(* IEC 61131-3 sources: PLC-IsaVODE/PLC-IsaVODE/samples/plc-programs (part 3) *)

(* ---- 394-TOD_TO_STRING.ST ---- *)
FUNCTION HOUR:INT
	VAR_INPUT
		ITOD :	UDINT;
	END_VAR
	hour := UDINT_TO_INT(itod / UDINT#3600000);
END_FUNCTION

FUNCTION MINUTE:INT

	VAR_INPUT
		ITOD :	UDINT;
	END_VAR

	minute := UDINT_TO_INT((itod / UDINT#60000) - ((itod / UDINT#3600000) * UDINT#60));

END_FUNCTION

FUNCTION_BLOCK TOD_TO_STRING_Block
	VAR_INPUT
		ITOD :	UDINT;
	END_VAR

	VAR_OUTPUT
		TOD_STRING :	STRING;
	END_VAR

	VAR
		st_tmp1 :	STRING;
		st_tmp2 :	STRING;
		cur_hours :	INT;
	END_VAR

	cur_hours := hour(ITOD);
	IF cur_hours = 0 THEN
	st_tmp2 := '%01dh';
	ELSE
	st_tmp2 := '%dh';
	END_IF;

	st_tmp1 := CONCAT(INT_TO_STRING(cur_hours),INT_TO_STRING(minute(ITOD)));
	TOD_STRING := CONCAT(st_tmp1,UDINT_TO_STRING(ITOD MOD UDINT#60000 / UDINT#1000));
END_FUNCTION_BLOCK

PROGRAM program0
  VAR
    LocalVar0 : UDINT;
	LocalOUT  : STRING;
	func_block : TOD_TO_STRING_Block;
  END_VAR
	func_block.ITOD  := LocalVar0;
	func_block();
	LocalOUT := func_block.TOD_STRING;
END_PROGRAM

CONFIGURATION Config0
  RESOURCE Res0 ON PLC
    TASK task0(INTERVAL := T#20ms,PRIORITY := 0);
    PROGRAM instance0 WITH task0 : program0;
  END_RESOURCE
END_CONFIGURATION

(* ---- 396-CLICK_MODE.ST ---- *)
FUNCTION_BLOCK CLICK_MODE_Block

	VAR_INPUT
		IN :	BOOL;
		T_LONG :	TIME := T#500ms;
	END_VAR

	VAR_OUTPUT
		LONG    :   BOOL;
		SINGLE_  :	BOOL;
		DOUBLE  :	BOOL;
		TP_LONG :	BOOL;
	END_VAR

	VAR
		Timer :	TP;
		cnt :	INT;
		last :	BOOL;
	END_VAR

	timer(in := IN, PT := T_LONG);
	single := FALSE;
	double := FALSE;

	IF timer.Q THEN
		IF NOT in AND last THEN	cnt := cnt + 1; END_IF;
	ELSE
		CASE cnt OF
			1 : single := TRUE;
			2 : double := TRUE;
		END_CASE;
		cnt := 0;
	END_IF;
	last := in;
	TP_LONG := NOT timer.Q AND (NOT LONG) AND IN;
	LONG := NOT timer.Q AND in;

END_FUNCTION_BLOCK

PROGRAM program0
	VAR
		IN :	BOOL;
		T_LONG :	TIME := T#500ms;
		SINGLE_ :	BOOL;
		DOUBLE :	BOOL;
		LONG :	BOOL;
		TP_LONG :	BOOL;

		func_block : CLICK_MODE_Block;
	END_VAR
	func_block.IN := IN;
	func_block.T_LONG := T_LONG;

	func_block();
	SINGLE_  := func_block.SINGLE_;
	DOUBLE  := func_block.DOUBLE;
	LONG  := func_block.LONG;
	TP_LONG  := func_block.TP_LONG;
END_PROGRAM

CONFIGURATION Config0
	RESOURCE Res0 ON PLC
		TASK task0(INTERVAL := T#20ms,PRIORITY := 0);
		PROGRAM instance0 WITH task0 : program0;
	END_RESOURCE
END_CONFIGURATION

(* ---- 397-IP4_TO_STRING.ST ---- *)
TYPE
  oscat_STRING10             : STRING;
END_TYPE

FUNCTION _BYTE_TO_INT:INT
	VAR_INPUT
		IN :	BYTE;
	END_VAR

	_BYTE_TO_INT := USINT_TO_INT(BYTE_TO_USINT(IN));
END_FUNCTION

FUNCTION BYTE_OF_DWORD:BYTE
	VAR_INPUT
		IN :	DWORD;
		N :	BYTE;
	END_VAR
	BYTE_OF_DWORD := DWORD_TO_BYTE(SHR(in,_BYTE_TO_INT(SHL(n,3))));
END_FUNCTION

FUNCTION_BLOCK IP4_TO_STRING_Block

	VAR_INPUT
		IP4 :	DWORD;
	END_VAR

	VAR_OUTPUT
		IP4_TO_STRING :	STRING;
	END_VAR

	VAR
		s1 :	oscat_string10;
		s2 :	oscat_string10;
	END_VAR

	s1 := CONCAT(BYTE_TO_STRING(BYTE_OF_DWORD(IP4,BYTE#1)),BYTE_TO_STRING(BYTE_OF_DWORD(IP4,BYTE#0)));
	s2 := CONCAT(BYTE_TO_STRING(BYTE_OF_DWORD(IP4,BYTE#3)),BYTE_TO_STRING(BYTE_OF_DWORD(IP4,BYTE#2)));
	IP4_TO_STRING := CONCAT(s2,s1);

END_FUNCTION_BLOCK

PROGRAM program0
	VAR
		IP4 :	DWORD;
		IP4_TO_STRING :	STRING;

		func_block : IP4_TO_STRING_Block;
	END_VAR
	func_block.IP4 := IP4;

	func_block();
	IP4_TO_STRING  := func_block.IP4_TO_STRING;
END_PROGRAM

CONFIGURATION Config0

  	RESOURCE Res0 ON PLC
    	TASK task0(INTERVAL := T#20ms,PRIORITY := 0);
    	PROGRAM instance0 WITH task0 : program0;
  	END_RESOURCE

END_CONFIGURATION

(* ---- 398-SHR_4UDE.ST ---- *)
FUNCTION_BLOCK SHR_4UDE_Block

	VAR_INPUT
		SET :	BOOL;
		D0 :	BOOL;
		D3 :	BOOL;
		CLK :	BOOL;
		DN :	BOOL;
		RST :	BOOL;
	END_VAR

	VAR_OUTPUT
		Q0 :	BOOL;
		Q1 :	BOOL;
		Q2 :	BOOL;
		Q3 :	BOOL;
	END_VAR

	VAR
		trig :	R_TRIG;
	END_VAR

	trig(clk := clk);

	IF set OR rst THEN
		Q0 := NOT RST;
		Q1 := Q0;
		Q2 := Q0;
		Q3 := Q0;
	ELSIF trig.Q THEN
		IF dn THEN
			Q0 := Q1;
			Q1 := Q2;
			Q2 := Q3;
			Q3 := D3;
		ELSE
			Q3 := Q2;
			Q2 := Q1;
			Q1 := Q0;
			Q0 := D0;
		END_IF;
	END_IF;

END_FUNCTION_BLOCK

PROGRAM program0

	VAR
		SET :	BOOL;
		D0 :	BOOL;
		D3 :	BOOL;
		CLK :	BOOL;
		DN :	BOOL;
		RST :	BOOL;
		Q0 :	BOOL;
		Q1 :	BOOL;
		Q2 :	BOOL;
		Q3 :	BOOL;
		func_block : SHR_4UDE_Block;
	END_VAR
	func_block.SET  :=SET;
	func_block.D0  :=D0;
	func_block.D3  :=D3;
	func_block.CLK  :=CLK;
	func_block.DN  :=DN;
	func_block.RST  :=RST;
	func_block();
	Q0 := func_block.Q0;
	Q1 := func_block.Q1;
	Q2 := func_block.Q2;
	Q3 := func_block.Q3;

END_PROGRAM

CONFIGURATION Config0
	RESOURCE Res0 ON PLC
		TASK task0(INTERVAL := T#20ms,PRIORITY := 0);
		PROGRAM instance0 WITH task0 : program0;
	END_RESOURCE
END_CONFIGURATION

(* ---- 399-MANUAL_1.ST ---- *)
FUNCTION_BLOCK MANUAL_1_Block

	VAR_INPUT
		_IN :	BOOL;
		MAN :	BOOL;
		M_I :	BOOL;
		SET :	BOOL;
		RST :	BOOL;
	END_VAR

	VAR_OUTPUT
		Q :	BOOL;
		STATUS :	BYTE;
	END_VAR

	VAR
		S_edge :	BOOL;
		_r_edge :	BOOL;
		edge :	BOOL;
	END_VAR

	IF NOT man THEN
		Q := _IN;
		STATUS := BYTE#100;
		edge := FALSE;
	ELSIF NOT s_edge AND set THEN
		Q := TRUE;
		edge := TRUE;
		status := BYTE#101;
	ELSIF NOT _r_edge AND rst THEN
		Q := FALSE;
		edge := TRUE;
		status := BYTE#102;
	ELSIF NOT edge THEN
		Q := M_I;
		status := BYTE#103;
	END_IF;

	(* remember levels of manual signals *)
	s_edge := SET;
	_r_edge := RST;

END_FUNCTION_BLOCK

PROGRAM program0

	VAR
		_IN :	BOOL;
		MAN :	BOOL;
		M_I :	BOOL;
		SET :	BOOL;
		RST :	BOOL;

		Q :	BOOL;
		STATUS :	BYTE;

		func_block : MANUAL_1_Block;
	END_VAR
	func_block._IN := _IN;
	func_block.MAN := MAN;
	func_block.M_I := M_I;
	func_block.SET := SET;
	func_block.RST := RST;
	func_block();
	Q := func_block.Q;
	STATUS := func_block.STATUS;

END_PROGRAM

CONFIGURATION Config0

	RESOURCE Res0 ON PLC
		TASK task0(INTERVAL := T#20ms,PRIORITY := 0);
		PROGRAM instance0 WITH task0 : program0;
	END_RESOURCE

END_CONFIGURATION

(* ---- 4-COUNT_CHAR.ST ---- *)
FUNCTION_BLOCK COUNT_CHAR
	VAR_INPUT
		STR :	STRING;
		CHR :	BYTE;
	END_VAR

	VAR_OUTPUT
		COUNT_CHAR :	INT;
	END_VAR

	VAR
		I :	INT;
		pos :	INT;
	END_VAR

	I := LEN(str);
	COUNT_CHAR := 0;
	FOR pos := 1 TO I DO
		IF INT_TO_BYTE(GET_CHAR(str,pos)) = CHR THEN COUNT_CHAR := COUNT_CHAR + 1; END_IF;
	END_FOR;
END_FUNCTION_BLOCK

(* ---- 401-STRING_TO_BUFFER.ST ---- *)
TYPE
	oscat_STRING250             : STRING(250);
	oscat_arb_0_249 			  : ARRAY [0..249] 	OF BYTE;
END_TYPE

FUNCTION_BLOCK _STRING_TO_BUFFER_Block
	VAR_INPUT
		STR :	oscat_STRING250;
		POS :	INT;
		SIZE :	UINT;
	END_VAR

	VAR_OUTPUT
		_STRING_TO_BUFFER :	INT;
	END_VAR

	VAR_IN_OUT
		PT :	oscat_arb_0_249;
	END_VAR

	VAR
		i :	INT;
		end :	INT;
		x :	INT;
	END_VAR

	IF pos < 0 THEN RETURN; END_IF;
	end := MIN(pos + LEN(str), UINT_TO_INT(size)) - 1;
	x:= 1;
	FOR i := pos TO end DO
		pt[i] := INT_TO_BYTE(GET_CHAR(str,x));
		x := x + 1;
	END_FOR;

	_STRING_TO_BUFFER := i;
END_FUNCTION_BLOCK

PROGRAM program0
	VAR
	    LocalVar1 : oscat_STRING250;
        LocalVar2 : INT;
        LocalVar3 : UINT;
		LocalInOut : oscat_arb_0_249;
		LocalOUT  : INT;
		func_block : _STRING_TO_BUFFER_Block;
  	END_VAR
	func_block.STR := LocalVar1;
    func_block.POS := LocalVar2;
    func_block.SIZE := LocalVar3;
	func_block.PT := LocalInOut;
	func_block();
	LocalOUT := func_block._STRING_TO_BUFFER;
	LocalInOut := func_block.PT;
END_PROGRAM

CONFIGURATION Config0
  	RESOURCE Res0 ON PLC
    	TASK task0(INTERVAL := T#20ms,PRIORITY := 0);
    	PROGRAM instance0 WITH task0 : program0;
  	END_RESOURCE
END_CONFIGURATION

(* ---- 402-SEL2_OF_3.ST ---- *)
FUNCTION_BLOCK SEL2_OF_3_Block

	VAR_INPUT
		IN1 :	REAL;
		IN2 :	REAL;
		IN3 :	REAL;
		D :	REAL;
	END_VAR

	VAR_OUTPUT
		Y :	REAL;
		W :	INT;
		E :	BOOL;
	END_VAR

	VAR
		D12 :	BOOL;
		D23 :	BOOL;
		D31 :	BOOL;
	END_VAR

	D12 := ABS(IN1-IN2) <= D;
	D23 := ABS(IN2-IN3) <= D;
	D31 := ABS(IN3-IN1) <= D;

	IF (D12 AND D23) OR (D12 AND D31) OR (D23 AND D31) THEN
		Y := (IN1 + IN2 + IN3) * 0.333333333333;
		E := FALSE;
		W := 0;
	ELSIF D12 THEN
		Y := (In1 + IN2) * 0.5;
		E := FALSE;
		W := 3;
	ELSIF D23 THEN
		Y := (In2 + IN3) * 0.5;
		E := FALSE;
		W := 1;
	ELSIF D31 THEN
		Y := (In3 + IN1) * 0.5;
		E := FALSE;
		W := 2;
	ELSE
		E := TRUE;
		W := 4;
	END_IF;

END_FUNCTION_BLOCK

PROGRAM program0

	VAR
		IN1 :	REAL;
		IN2 :	REAL;
		IN3 :	REAL;
		D :	REAL;
		Y :	REAL;
		W :	INT;
		E :	BOOL;
		func_block : SEL2_OF_3_Block;
  	END_VAR
	func_block.IN1  :=IN1;
	func_block.IN2  :=IN2;
	func_block.IN3  :=IN3;
	func_block.D  :=D;
	func_block();
	Y := func_block.Y;
	W := func_block.W;
	E := func_block.E;

END_PROGRAM

CONFIGURATION Config0

	RESOURCE Res0 ON PLC
		TASK task0(INTERVAL := T#20ms,PRIORITY := 0);
		PROGRAM instance0 WITH task0 : program0;
	END_RESOURCE

END_CONFIGURATION

(* ---- 403-CLOG.ST ---- *)
TYPE oscat_complex :
  STRUCT
	re : REAL;
	im : REAL;
  END_STRUCT;
END_TYPE

FUNCTION ATAN2:REAL
	VAR_INPUT
		X :	REAL;
		Y :	REAL;
	END_VAR

	IF X > 0.0 THEN
		ATAN2 := ATAN(Y/X);
	ELSIF X < 0.0 THEN
		IF Y >= 0.0 THEN
			ATAN2 := ATAN(Y/X) + 3.14159265358979323846264338327950288;
		ELSE
			ATAN2 := ATAN(Y/X) - 3.14159265358979323846264338327950288;
		END_IF;
	ELSIF Y > 0.0 THEN
		ATAN2 := 1.5707963267948965580;
	ELSIF Y < 0.0 THEN
		ATAN2 := -1.5707963267948965580;
	ELSE
		ATAN2 := 0.0;
	END_IF;

END_FUNCTION

FUNCTION HYPOT:REAL
	VAR_INPUT
		X :	REAL;
		Y :	REAL;
	END_VAR

	HYPOT := SQRT(x*x + y*y);
END_FUNCTION

FUNCTION_BLOCK CLOG_Block

	VAR_INPUT
		X :	oscat_complex;
	END_VAR

	VAR_OUTPUT
		CLOG :	oscat_complex;
	END_VAR

	CLOG.re := LN(HYPOT(X.re, X.im));
	CLOG.im := ATAN2(X.im, X.re);

END_FUNCTION_BLOCK

PROGRAM program0
  VAR
    LocalVar0 : oscat_complex;
	LocalOUT  : oscat_complex;
	func_block : CLOG_Block;
  END_VAR
	func_block.X  := LocalVar0;
	func_block();
	LocalOUT := func_block.CLOG;
END_PROGRAM

CONFIGURATION Config0
  RESOURCE Res0 ON PLC
    TASK task0(INTERVAL := T#20ms,PRIORITY := 0);
    PROGRAM instance0 WITH task0 : program0;
  END_RESOURCE
END_CONFIGURATION

(* ---- 406-ELEMENT_GET.ST ---- *)
TYPE
	oscat_STRING250             : STRING;
END_TYPE

FUNCTION_BLOCK ELEMENT_GET_Block

	VAR_INPUT
		SEP :	BYTE;
		POS :	INT;
	END_VAR

	VAR_IN_OUT
		ELEMENT :	oscat_STRING250;
	END_VAR

	VAR_OUTPUT
		ELEMENT_GET :	oscat_STRING250;
	END_VAR

	VAR
		i :	INT;
		i2 :	INT;
		cnt :	INT;
		size :	INT;
	END_VAR

	cnt := 0;
	size := LEN(ELEMENT);

	FOR i := 1 TO size DO
		IF cnt = POS THEN EXIT; END_IF;
		IF INT_TO_BYTE(GET_CHAR(ELEMENT,i)) = SEP THEN cnt := cnt + 1; END_IF;
	END_FOR;

	FOR i2 := i TO size DO
		IF INT_TO_BYTE(GET_CHAR(ELEMENT,i2)) = SEP THEN EXIT; END_IF;
	END_FOR;

	IF i2 > i THEN
		ELEMENT_GET := MID(ELEMENT,i2-i,i);
	ELSE
		ELEMENT_GET := '';
	END_IF;

END_FUNCTION_BLOCK

PROGRAM program0
	VAR
		SEP :	BYTE;
		POS :	INT;
		ELEMENT :	oscat_STRING250;
		ELEMENT_GET :	oscat_STRING250;

		func_block : ELEMENT_GET_Block;
	END_VAR
	func_block.SEP    :=SEP    ;
	func_block.POS:=POS;
	func_block.ELEMENT     :=ELEMENT     ;
	func_block();
	ELEMENT    := func_block.ELEMENT    ;
	ELEMENT_GET:= func_block.ELEMENT_GET;

END_PROGRAM

CONFIGURATION Config0
  RESOURCE Res0 ON PLC
    TASK task0(INTERVAL := T#20ms,PRIORITY := 0);
    PROGRAM instance0 WITH task0 : program0;
  END_RESOURCE
END_CONFIGURATION

(* ---- 407-FILTER_MAV_DW.ST ---- *)
TYPE
  oscat_ardw_0_31             : ARRAY [0..31]   OF DWORD;
END_TYPE

FUNCTION INC1:INT

	VAR_INPUT
		X :	INT;
		N :	INT;
	END_VAR

	IF X >= N - 1 THEN
		INC1 := 0;
	ELSE
		INC1 := X + 1;
	END_IF;
END_FUNCTION

FUNCTION_BLOCK FILTER_MAV_DW

	VAR_INPUT
		X :	DWORD;
		N :	UINT;
		RST :	BOOL;
	END_VAR

	VAR_OUTPUT
		Y :	DWORD;
	END_VAR

	VAR
		init :	BOOL;
		buffer :	oscat_ardw_0_31;
		i :	INT;
		tmp :	INT;
	END_VAR

	N := MIN(N, UINT#32);

	(* startup initialisation *)
	IF NOT init OR rst OR N = UINT#0 THEN
		init := TRUE;
		tmp := UINT_TO_INT(N)-1;
		FOR i := 0 TO tmp DO
			buffer[i] := X;
		END_FOR;
		Y := X;
	ELSE
		tmp := UINT_TO_INT(N);
		i := INC1(i, tmp);
		Y := UDINT_TO_DWORD(DWORD_TO_UDINT(Y) + (DWORD_TO_UDINT(X) - DWORD_TO_UDINT(buffer[i])) / UINT_TO_UDINT(N));
		buffer[i] := X;
	END_IF;

END_FUNCTION_BLOCK

PROGRAM program0
  VAR
	X :	DWORD;
	N :	UINT;
	RST :	BOOL;

	Y :	DWORD;

	func_block : FILTER_MAV_DW;
  END_VAR
	func_block.X  := X;
	func_block.N  := N;
	func_block.RST  := RST;
	func_block();
	Y := func_block.Y;
END_PROGRAM

CONFIGURATION Config0

	RESOURCE Res0 ON PLC
		TASK task0(INTERVAL := T#20ms,PRIORITY := 0);
		PROGRAM instance0 WITH task0 : program0;
	END_RESOURCE
END_CONFIGURATION

(* ---- 409-STATUS_TO_ESR.ST ---- *)
TYPE
  oscat_esr_collect_data      : ARRAY [0..7]    OF BYTE;
END_TYPE

TYPE oscat_esr_data :
  STRUCT
	typ    : BYTE;
	adress : STRING;
	DS     : UDINT;
	TS     : TIME;
	data   : oscat_esr_collect_data;
  END_STRUCT;
END_TYPE

FUNCTION_BLOCK STATUS_TO_ESR_Block

	VAR_INPUT
		STATUS :	BYTE;
		ADRESS :	STRING;
		DT_IN :	UDINT;
		TS :	TIME;
	END_VAR

	VAR_OUTPUT
		STATUS_TO_ESR :	oscat_esr_data;
	END_VAR

	IF status < BYTE#100 THEN
		status_to_ESR.typ := BYTE#1;
	ELSIF status < BYTE#200 THEN
		status_to_ESR.typ := BYTE#2;
	ELSE
		status_to_ESR.typ := BYTE#3;
	END_IF;
	status_to_ESR.adress:= adress;
	status_to_ESR.DS := DT_in;
	status_to_ESR.TS := TS;
	status_to_ESR.data[0] := status;
END_FUNCTION_BLOCK

PROGRAM program0
	VAR
		STATUS :	BYTE;
		ADRESS :	STRING;
		DT_IN  :	UDINT;
		TS     :	TIME;
		STATUS_TO_ESR :	oscat_esr_data;

		func_block : STATUS_TO_ESR_Block;
	END_VAR
	func_block.STATUS := STATUS;
	func_block.ADRESS := ADRESS;
	func_block.DT_IN := DT_IN ;
	func_block.TS    := TS    ;

	func_block();
	STATUS_TO_ESR  := func_block.STATUS_TO_ESR;
END_PROGRAM

CONFIGURATION Config0
	RESOURCE Res0 ON PLC
		TASK task0(INTERVAL := T#20ms,PRIORITY := 0);
		PROGRAM instance0 WITH task0 : program0;
	END_RESOURCE
END_CONFIGURATION

(* ---- 410-V3_PAR.ST ---- *)
TYPE oscat_vector_3:
	STRUCT
		X : REAL;
		Y : REAL;
		Z : REAL;
	END_STRUCT;
END_TYPE

FUNCTION_BLOCK V3_ABS_Block

	VAR_INPUT
		A :	oscat_vector_3;
	END_VAR

	VAR_OUTPUT
		V3_ABS :	REAL;
	END_VAR

	V3_ABS := SQRT(A.X * A.X + A.Y * A.Y + A.Z * A.Z);

END_FUNCTION_BLOCK

FUNCTION_BLOCK V3_XPRO_Block
	VAR_INPUT
		A :	oscat_vector_3;
		B :	oscat_vector_3;
	END_VAR

	VAR_OUTPUT
		V3_XPRO :	oscat_vector_3;
	END_VAR

	V3_XPRO.X := A.Y * B.Z - A.Z * B.Y;
	V3_XPRO.Y := A.Z * B.X - A.X * B.Z;
	V3_XPRO.Z := A.X * B.Y - A.Y * B.X;

END_FUNCTION_BLOCK

FUNCTION_BLOCK V3_PAR_Block
	VAR_INPUT
		A :	oscat_vector_3;
		B :	oscat_vector_3;
	END_VAR

	VAR_OUTPUT
		V3_PAR :	BOOL;
	END_VAR

	VAR
		V3_XPRO :	V3_XPRO_Block;
		V3_ABS :	V3_ABS_Block;
	END_VAR

	V3_XPRO(A:=A,B:=B);
	V3_ABS(A:=V3_XPRO.V3_XPRO);

	V3_PAR := V3_ABS.V3_ABS = 0.0;

END_FUNCTION_BLOCK

PROGRAM program0
  	VAR
		A :	oscat_vector_3;
		B :	oscat_vector_3;
		V3_PAR :	BOOL;
		func_block : V3_PAR_Block;
  	END_VAR
	func_block.A := A;
	func_block.B := B;
	func_block();
	V3_PAR := func_block.V3_PAR;
END_PROGRAM

CONFIGURATION Config0
  RESOURCE Res0 ON PLC
    TASK task0(INTERVAL := T#20ms,PRIORITY := 0);
    PROGRAM instance0 WITH task0 : program0;
  END_RESOURCE
END_CONFIGURATION

(* ---- 411-FILTER_WAV.ST ---- *)
TYPE
  oscat_arr_0_15              : ARRAY [0..15]   OF REAL;
END_TYPE

FUNCTION INC1:INT

	VAR_INPUT
		X :	INT;
		N :	INT;
	END_VAR

	IF X >= N - 1 THEN
		INC1 := 0;
	ELSE
		INC1 := X + 1;
	END_IF;
END_FUNCTION

FUNCTION DEC1:INT

	VAR_INPUT
		X :	INT;
		N :	INT;
	END_VAR

	IF X = 0 THEN
		DEC1 := N - 1;
	ELSE
		DEC1 := X - 1;
	END_IF;

END_FUNCTION

FUNCTION_BLOCK FILTER_WAV
	VAR_INPUT
		X :	REAL;
		W :	oscat_arr_0_15;
		RST :	BOOL;
	END_VAR

	VAR_OUTPUT
		Y :	REAL;
	END_VAR

	VAR
		init :	BOOL;
		buffer :	oscat_arr_0_15;
		i :	INT;
		n :	INT;
	END_VAR

	IF NOT init OR rst THEN
		init := TRUE;
		FOR i := 0 TO 15 DO
			buffer[i] := X;
		END_FOR;
		i := 15;
		Y := X;
	ELSE
		i := INC1(i, 16);
		buffer[i] := X;
	END_IF;

	Y := 0.0;
	FOR n := 0 TO 15 DO
		Y := buffer[i] * W[n] + Y;
		i := DEC1(i, 16);
	END_FOR;
END_FUNCTION_BLOCK

PROGRAM program0
  VAR
	X :	REAL;
	W :	oscat_arr_0_15;
	RST :	BOOL;

	Y :	REAL;

	func_block : FILTER_WAV;
  END_VAR
	func_block.X  := X;
	func_block.W  := W;
	func_block.RST  := RST;
	func_block();
	Y := func_block.Y;
END_PROGRAM

CONFIGURATION Config0

	RESOURCE Res0 ON PLC
		TASK task0(INTERVAL := T#20ms,PRIORITY := 0);
		PROGRAM instance0 WITH task0 : program0;
	END_RESOURCE
END_CONFIGURATION

(* ---- 412-STRING_TO_TOD.ST ---- *)
FUNCTION_BLOCK STRING_TO_TOD_Block

  VAR_INPUT
    _TOD :	STRING;
  END_VAR

  VAR_OUTPUT
    out_STRING_TO_TOD :	UDINT;
  END_VAR

  VAR
    pos :	INT;
    i :	INT;
    tmp :	STRING;
    tmp2 :	STRING;
  END_VAR

  out_STRING_TO_TOD := UDINT#0;
  i := LEN(_TOD);
  pos :=FIND(_TOD,'#');

  IF pos>0 AND i>pos THEN
    tmp := RIGHT(_TOD,LEN(_TOD)-pos);
    pos := FIND(tmp,':');
    IF pos>1 THEN
      tmp2 := LEFT(tmp,pos-1);
      tmp := RIGHT(tmp,LEN(tmp)-pos);
      out_STRING_TO_TOD := STRING_TO_UDINT(tmp2) * UDINT#3600000;

      pos :=FIND(tmp,':');
      IF pos>1 THEN
        tmp2 := LEFT(tmp,pos-1);
        tmp := RIGHT(tmp,LEN(tmp)-pos);
        out_STRING_TO_TOD := out_STRING_TO_TOD + STRING_TO_UDINT(tmp2) * UDINT#60000;

        out_STRING_TO_TOD := out_STRING_TO_TOD + STRING_TO_UDINT(tmp) * UDINT#1000;
      END_IF;
    END_IF;
  END_IF;

END_FUNCTION_BLOCK

PROGRAM program0
  VAR
    _TOD :	STRING;
  	out_STRING_TO_TOD :	UDINT;
    func_block : STRING_TO_TOD_Block;
  END_VAR
	func_block._TOD  := _TOD;
	func_block();
	out_STRING_TO_TOD  := func_block.out_STRING_TO_TOD;
END_PROGRAM

CONFIGURATION Config0
	RESOURCE Res0 ON PLC
		TASK task0(INTERVAL := T#20ms,PRIORITY := 0);
		PROGRAM instance0 WITH task0 : program0;
	END_RESOURCE
END_CONFIGURATION

(* ---- 414-SETUP_WEEKDAYS2.ST ---- *)
TYPE
  oscat_ELEMENT_WEEKDAYS2	: ARRAY [1..7] OF STRING;
  oscat_WEEKDAYS2			: ARRAY [1..3]  OF oscat_ELEMENT_WEEKDAYS2 := [0, 0, 0];
END_TYPE

FUNCTION_BLOCK SETUP_WEEKDAYS2_Block

	VAR_IN_OUT
		WEEKDAYS2 :	oscat_WEEKDAYS2;
	END_VAR

	VAR
		init :	BOOL;
	END_VAR

	IF init THEN RETURN; END_IF;
	init := TRUE;

	WEEKDAYS2[1][01] := 'Mo';
	WEEKDAYS2[1][02] := 'Tu';
	WEEKDAYS2[1][03] := 'We';
	WEEKDAYS2[1][04] := 'Th';
	WEEKDAYS2[1][05] := 'Fr';
	WEEKDAYS2[1][06] := 'Sa';
	WEEKDAYS2[1][07] := 'Su';

	WEEKDAYS2[2][01] := 'Mo';
	WEEKDAYS2[2][02] := 'Di';
	WEEKDAYS2[2][03] := 'Mi';
	WEEKDAYS2[2][04] := 'Do';
	WEEKDAYS2[2][05] := 'Fr';
	WEEKDAYS2[2][06] := 'Sa';
	WEEKDAYS2[2][07] := 'So';

	WEEKDAYS2[3][01] := 'Lu';
	WEEKDAYS2[3][02] := 'Ma';
	WEEKDAYS2[3][03] := 'Me';
	WEEKDAYS2[3][04] := 'Je';
	WEEKDAYS2[3][05] := 'Ve';
	WEEKDAYS2[3][06] := 'Sa';
	WEEKDAYS2[3][07] := 'Di';
END_FUNCTION_BLOCK

PROGRAM program0

	VAR
		WEEKDAYS2 :	oscat_WEEKDAYS2;
		func_block : SETUP_WEEKDAYS2_Block;
	END_VAR
		func_block.WEEKDAYS2 :=WEEKDAYS2;
		func_block();
		WEEKDAYS2 := func_block.WEEKDAYS2;

END_PROGRAM

CONFIGURATION Config0

	RESOURCE Res0 ON PLC
		TASK task0(INTERVAL := T#20ms,PRIORITY := 0);
		PROGRAM instance0 WITH task0 : program0;
	END_RESOURCE

END_CONFIGURATION

(* ---- 415-STACK_16.ST ---- *)
TYPE
  oscat_ardw_0_15             : ARRAY [0..15]   OF DWORD;
END_TYPE

FUNCTION_BLOCK STACK_16_Block

	VAR_INPUT
		DIN :	DWORD;
		E :	BOOL := TRUE;
		RD :	BOOL;
		WD :	BOOL;
		RST :	BOOL;
	END_VAR

	VAR_OUTPUT
		DOUT :	DWORD;
		EMPTY :	BOOL := TRUE;
		FULL :	BOOL;
	END_VAR

	VAR
		pt :	INT;
		stack :	oscat_ardw_0_15;
	END_VAR

	IF RST THEN
		pt := 0;
		EMPTY := TRUE;
		FULL := FALSE;
		Dout := DWORD#0;
	ELSIF E THEN
		IF NOT EMPTY AND RD THEN
			pt := pt - 1;
			Dout := stack[pt];
			EMPTY := pt = 0;
			FULL := FALSE;
		END_IF;
		IF NOT FULL AND WD THEN
			stack[pt] := Din;
			pt := pt + 1;
			FULL := pt > 15;
			EMPTY := FALSE;
		END_IF;
	END_IF;

END_FUNCTION_BLOCK

PROGRAM program0
	VAR
		DIN :	DWORD;
		E :	BOOL := TRUE;
		RD :	BOOL;
		WD :	BOOL;
		RST :	BOOL;
		DOUT :	DWORD;
		EMPTY :	BOOL := TRUE;
		FULL :	BOOL;
		func_block : STACK_16_Block;
	END_VAR
		func_block.DIN  := DIN;
		func_block.E  := E;
		func_block.RD  := RD;
		func_block.WD  := WD;
		func_block.RST  := RST;
		func_block();
		DOUT := func_block.DOUT;
		EMPTY := func_block.EMPTY;
		FULL := func_block.FULL;

END_PROGRAM

CONFIGURATION Config0

	RESOURCE Res0 ON PLC
		TASK task0(INTERVAL := T#20ms,PRIORITY := 0);
		PROGRAM instance0 WITH task0 : program0;
	END_RESOURCE

END_CONFIGURATION

(* ---- 416-FILTER_MAV_W.ST ---- *)
TYPE
  oscat_FILTER_MAV_W          : ARRAY [0..31]   OF WORD;
END_TYPE

FUNCTION INC1:INT

	VAR_INPUT
		X :	INT;
		N :	INT;
	END_VAR

	IF X >= N - 1 THEN
		INC1 := 0;
	ELSE
		INC1 := X + 1;
	END_IF;
END_FUNCTION

FUNCTION_BLOCK FILTER_MAV_W
	VAR_INPUT
		X :	WORD;
		N :	UINT;
		RST :	BOOL;
	END_VAR

	VAR_OUTPUT
		Y :	WORD;
	END_VAR

	VAR
		init :	BOOL;
		buffer :	oscat_FILTER_MAV_W;
		i :	INT;
		sum :	UDINT;
		tmp :	INT;
	END_VAR

	N := MIN(N, UINT#32);

	(* startup initialisation *)
	IF NOT init OR rst OR N = UINT#0 THEN
		init := TRUE;
		tmp := UINT_TO_INT(N) - 1;
		FOR i := 1 TO tmp DO
			buffer[i] := X;
		END_FOR;
		sum := UINT_TO_UDINT(WORD_TO_UINT(Y) * N);
		Y := X;
	ELSE
		tmp := UINT_TO_INT(N);
		i := INC1(i, tmp);
		sum := sum + WORD_TO_UDINT(X) - WORD_TO_UDINT(buffer[i]);
		Y := UDINT_TO_WORD(sum / UINT_TO_UDINT(N));
		buffer[i] := X;
	END_IF;

END_FUNCTION_BLOCK

PROGRAM program0
  VAR
	X :	WORD;
	N :	UINT;
	RST :	BOOL;

	Y :	WORD;

	func_block : FILTER_MAV_W;
  END_VAR
	func_block.X  := X;
	func_block.N  := N;
	func_block.RST  := RST;
	func_block();
	Y := func_block.Y;
END_PROGRAM

CONFIGURATION Config0

	RESOURCE Res0 ON PLC
		TASK task0(INTERVAL := T#20ms,PRIORITY := 0);
		PROGRAM instance0 WITH task0 : program0;
	END_RESOURCE
END_CONFIGURATION

(* ---- 418-V3_NORM.ST ---- *)
TYPE oscat_vector_3:
	STRUCT
		X : REAL;
		Y : REAL;
		Z : REAL;
	END_STRUCT;
END_TYPE

FUNCTION_BLOCK V3_ABS_Block

	VAR_INPUT
		A :	oscat_vector_3;
	END_VAR

	VAR_OUTPUT
		V3_ABS :	REAL;
	END_VAR

	V3_ABS := SQRT(A.X * A.X + A.Y * A.Y + A.Z * A.Z);

END_FUNCTION_BLOCK

FUNCTION_BLOCK V3_SMUL_Block
	VAR_INPUT
		A :	oscat_vector_3;
		M :	REAL;
	END_VAR

	VAR_OUTPUT
		V3_SMUL :	oscat_vector_3;
	END_VAR

	V3_SMUL.X := A.X * M;
	V3_SMUL.Y := A.Y * M;
	V3_SMUL.Z := A.Z * M;
END_FUNCTION_BLOCK

FUNCTION_BLOCK V3_NORM_Block

	VAR_INPUT
		A :	oscat_vector_3;
	END_VAR

	VAR_OUTPUT
		V3_NORM :	oscat_vector_3;
	END_VAR

	VAR
		la :	REAL;
		V3_SMUL :	V3_SMUL_Block;
		V3_ABS :	V3_ABS_Block;
	END_VAR

	V3_ABS(A:=A);
	la:=V3_ABS.V3_ABS;

	IF la > 0.0 THEN
		V3_SMUL(A:=A,M:=1.0/la);
		V3_NORM:=V3_SMUL.V3_SMUL;
	ELSE
		V3_NORM.X := 0.0;
		V3_NORM.Y := 0.0;
		V3_NORM.Z := 0.0;
	END_IF;

END_FUNCTION_BLOCK

PROGRAM program0
  	VAR
		A :	oscat_vector_3;
		V3_NORM :	oscat_vector_3;
		func_block : V3_NORM_Block;
  	END_VAR
	func_block.A := A;
	func_block();
	V3_NORM := func_block.V3_NORM;
END_PROGRAM

CONFIGURATION Config0
  RESOURCE Res0 ON PLC
    TASK task0(INTERVAL := T#20ms,PRIORITY := 0);
    PROGRAM instance0 WITH task0 : program0;
  END_RESOURCE
END_CONFIGURATION

(* ---- 420-PRESSURE.ST ---- *)
FUNCTION_BLOCK PRESSURE_Block

	VAR_INPUT
		MWS :	REAL;
		TORR :	REAL;
		ATT :	REAL;
		ATM :	REAL;
		PA :	REAL;
		BAR :	REAL;
	END_VAR

	VAR_OUTPUT
		YMWS :	REAL;
		YTORR :	REAL;
		YATT :	REAL;
		YATM :	REAL;
		YPA :	REAL;
		YBAR :	REAL;
	END_VAR

	Ybar := bar +
			pa * 1.0E-5 +
			0.980665 * att +
			1.01325 * atm +
			0.001333224 * torr +
			0.0980665 * mws;
	Ymws := ybar * 10.1971621297793;
	Ytorr := ybar * 750.0615050434140;
	Yatt := ybar * 1.0197162129779;
	yatm := ybar * 0.9869232667160;
	Ypa := ybar * 100000.0;

END_FUNCTION_BLOCK

PROGRAM program0

	VAR
		MWS :	REAL;
		TORR :	REAL;
		ATT :	REAL;
		ATM :	REAL;
		PA :	REAL;
		BAR :	REAL;

		YMWS :	REAL;
		YTORR :	REAL;
		YATT :	REAL;
		YATM :	REAL;
		YPA :	REAL;
		YBAR :	REAL;
		func_block : PRESSURE_Block;
  	END_VAR
	func_block.MWS := MWS;
	func_block.TORR := TORR;
	func_block.ATT := ATT;
	func_block.ATM := ATM;
	func_block.PA := PA;
	func_block.BAR := BAR;
	func_block();
	YMWS := func_block.YMWS;
	YTORR := func_block.YTORR;
	YATT := func_block.YATT;
	YATM := func_block.YATM;
	YPA := func_block.YPA;
	YBAR := func_block.YBAR;

END_PROGRAM

CONFIGURATION Config0

  	RESOURCE Res0 ON PLC
    	TASK task0(INTERVAL := T#20ms,PRIORITY := 0);
    	PROGRAM instance0 WITH task0 : program0;
  	END_RESOURCE

END_CONFIGURATION

(* ---- 422-POLYNOM_INT.ST ---- *)
TYPE
	oscat_Polynom_ARRAY_X       : ARRAY [0..1]    OF REAL;
END_TYPE

TYPE
	oscat_Polynom_XY            : ARRAY [1..5]  OF oscat_Polynom_ARRAY_X := [0, 0, 0, 0, 0];
END_TYPE

FUNCTION_BLOCK POLYNOM_INT_Block

	VAR_INPUT
		X :	REAL;
		XY :	oscat_Polynom_XY;
	END_VAR

	VAR_INPUT
		PTS :	INT;
	END_VAR

	VAR_OUTPUT
		POLYNOM_INT :	REAL;
	END_VAR

	VAR
		XY2 :	oscat_Polynom_XY;
	END_VAR

	VAR
		I :	INT;
		J :	INT;
		J_1 :	INT;
		J_I :	INT;
		INIT :	BOOL;
	END_VAR

	pts := MIN_INT(pts, 5);

	IF (init = FALSE) THEN
		init := TRUE;

		FOR i := 1 TO pts DO
			FOR j := 0 TO 1 DO
					XY2[i][j] := XY[i][j];
			END_FOR;
		END_FOR;

		FOR i := 1 TO pts DO
			J := pts;
			WHILE (J >= i+1) DO
			j_i := j-i;
			j_1 := J-1;
			XY2[j][1] := (XY2[j][1] - XY2[j_1][1]) / (XY2[j][0] - XY2[j_i][0]);
			j := j - 1;
			END_WHILE;
		END_FOR;
	END_IF;

END_FUNCTION_BLOCK

PROGRAM program0

	VAR
		X :	REAL;
		XY :	oscat_Polynom_XY;
		PTS :	INT;

		OUT :	REAL;
		func_block : POLYNOM_INT_Block;
  	END_VAR

	func_block.X := X;
	func_block.XY := XY;
	func_block.PTS := PTS;
	func_block();
	OUT := func_block.POLYNOM_INT;

END_PROGRAM

CONFIGURATION Config0

  	RESOURCE Res0 ON PLC
    	TASK task0(INTERVAL := T#20ms,PRIORITY := 0);
    	PROGRAM instance0 WITH task0 : program0;
  	END_RESOURCE

END_CONFIGURATION

(* ---- 424-ARRAY_TREND.ST ---- *)
TYPE
	oscat_pt_ARRAY: ARRAY [1..100] OF REAL;
END_TYPE

FUNCTION BIT_OF_DWORD:BOOL
	VAR_INPUT
		IN :	DWORD;
		N :	INT;
	END_VAR
	BIT_OF_DWORD := (SHR(in,n) AND DWORD#1) > DWORD#0;
END_FUNCTION

FUNCTION EVEN:BOOL
	VAR_INPUT
		IN :	DINT;
	END_VAR
	even := NOT BIT_OF_DWORD(DINT_TO_DWORD(in),0);
END_FUNCTION

FUNCTION_BLOCK ARRAY_TREND_Block
	VAR_IN_OUT
		PT :	oscat_pt_ARRAY;
	END_VAR

	VAR_INPUT
		SIZE :	UINT;
	END_VAR

	VAR_OUTPUT
		ARRAY_TREND :	REAL;
	END_VAR

	VAR
		d :	INT;
		i :	INT;
		stop :	INT;
		stop2 :	INT;
		x :	REAL;
	END_VAR

	x := 0.0;
	stop :=LIMIT_INT(1,UINT_TO_INT(size),1000);
	stop2 := WORD_TO_INT(SHR(INT_TO_WORD(stop),1));
	IF even(INT_TO_DINT(stop)) THEN d:=0; ELSE d:=1;END_IF;

	FOR i := 1 TO stop2+d DO
		x := x - pt[i];
	END_FOR;
	FOR i := stop2+1 TO stop DO
		x := x + pt[i];
	END_FOR;
	array_trend := x / INT_TO_REAL(stop2+d);

END_FUNCTION_BLOCK

PROGRAM program0
  VAR
    LocalVar0 : oscat_pt_ARRAY;
    LocalVar1 : UINT;
	LocalOUT  : REAL;
	func_block : ARRAY_TREND_Block;
  END_VAR
	func_block.pt := LocalVar0;
	func_block.size := LocalVar1;
	func_block();
	LocalOUT := func_block.ARRAY_TREND;

END_PROGRAM

CONFIGURATION Config0
  RESOURCE Res0 ON PLC
    TASK task0(INTERVAL := T#20ms,PRIORITY := 0);
    PROGRAM instance0 WITH task0 : program0;
  END_RESOURCE
END_CONFIGURATION

(* ---- 425-SETUP_WEEKDAYS.ST ---- *)
TYPE
  oscat_ELEMENT_WEEKDAYS	: ARRAY [1..7] OF STRING;
  oscat_WEEKDAYS			: ARRAY [1..3]  OF oscat_ELEMENT_WEEKDAYS := [0, 0, 0];
END_TYPE

FUNCTION_BLOCK SETUP_WEEKDAYS

	VAR_IN_OUT
		WEEKDAYS :	oscat_WEEKDAYS;
	END_VAR

	VAR
		init :	BOOL;
	END_VAR

	IF init THEN RETURN; END_IF;
	init := TRUE;

	WEEKDAYS[1][01] := 'Monday';
	WEEKDAYS[1][02] := 'Tuesday';
	WEEKDAYS[1][03] := 'Wednesday';
	WEEKDAYS[1][04] := 'Thursday';
	WEEKDAYS[1][05] := 'Friday';
	WEEKDAYS[1][06] := 'Saturday';
	WEEKDAYS[1][07] := 'Sunday';

	WEEKDAYS[2][01] := 'Montag';
	WEEKDAYS[2][02] := 'Dienstag';
	WEEKDAYS[2][03] := 'Mittwoch';
	WEEKDAYS[2][04] := 'Donnerstag';
	WEEKDAYS[2][05] := 'Freitag';
	WEEKDAYS[2][06] := 'Samstag';
	WEEKDAYS[2][07] := 'Sonntag';

	WEEKDAYS[3][01] := 'Lundi';
	WEEKDAYS[3][02] := 'Mardi';
	WEEKDAYS[3][03] := 'Mercredi';
	WEEKDAYS[3][04] := 'Jeudi';
	WEEKDAYS[3][05] := 'Vendredi';
	WEEKDAYS[3][06] := 'Samedi';
	WEEKDAYS[3][07] := 'Dimanche';
END_FUNCTION_BLOCK

PROGRAM program0
  VAR
    WEEKDAYS :	oscat_WEEKDAYS;
	func_block : SETUP_WEEKDAYS;
  END_VAR
	func_block.WEEKDAYS  := WEEKDAYS;
	func_block();
	WEEKDAYS := func_block.WEEKDAYS;

END_PROGRAM

CONFIGURATION Config0
  RESOURCE Res0 ON PLC
    TASK task0(INTERVAL := T#20ms,PRIORITY := 0);
    PROGRAM instance0 WITH task0 : program0;
  END_RESOURCE
END_CONFIGURATION

(* ---- 426-V3_ANG.ST ---- *)
TYPE oscat_vector_3:
	STRUCT
		X : REAL;
		Y : REAL;
		Z : REAL;
	END_STRUCT;
END_TYPE

FUNCTION_BLOCK V3_ABS_Block
	VAR_INPUT
		A :	oscat_vector_3;
	END_VAR

	VAR_OUTPUT
		V3_ABS : REAL;
	END_VAR

	V3_ABS := SQRT(A.X * A.X + A.Y * A.Y + A.Z * A.Z);

END_FUNCTION_BLOCK

FUNCTION_BLOCK V3_DPRO_Block

	VAR_INPUT
		A :	oscat_vector_3;
		B :	oscat_vector_3;
	END_VAR

	VAR_OUTPUT
		V3_DPRO :	REAL;
	END_VAR

	V3_DPRO := A.X * B.X + A.Y * B.Y + A.Z * B.Z;

END_FUNCTION_BLOCK

FUNCTION_BLOCK V3_ANG_Block

	VAR_INPUT
		A :	oscat_vector_3;
		B :	oscat_vector_3;
	END_VAR

	VAR_OUTPUT
		V3_ANG :	REAL;
	END_VAR

	VAR
		d :	REAL;
		V3_ABS :	V3_ABS_Block;
		V3_DPRO :	V3_DPRO_Block;
	END_VAR

	V3_ABS(A:=A);
	d :=V3_ABS.V3_ABS;

	V3_ABS(A:=B);
	d := d * V3_ABS.V3_ABS;

	IF d > 0.0 THEN
		V3_DPRO(A:=A,B:=B);
		V3_ANG := ACOS(LIMIT(-1.0, V3_DPRO.V3_DPRO / d,1.0));
	ELSE
		V3_ANG := 0.0;

	END_IF;

END_FUNCTION_BLOCK

PROGRAM program0
  	VAR
		A :	oscat_vector_3;
		B :	oscat_vector_3;
		V3_ANG :	REAL;
		func_block : V3_ANG_Block;
  	END_VAR
	func_block.A := A;
	func_block.B := B;
	func_block();
	V3_ANG := func_block.V3_ANG;
END_PROGRAM

CONFIGURATION Config0
  RESOURCE Res0 ON PLC
    TASK task0(INTERVAL := T#20ms,PRIORITY := 0);
    PROGRAM instance0 WITH task0 : program0;
  END_RESOURCE
END_CONFIGURATION

(* ---- 427-FILL.ST ---- *)
FUNCTION_BLOCK CHR_TO_STRING_Block
	VAR_INPUT
		C :	BYTE;
	END_VAR

	VAR_OUTPUT
		CHR_TO_STRING :	STRING;
	END_VAR

	CHR_TO_STRING := BYTE_TO_STRING(C);

END_FUNCTION_BLOCK

FUNCTION BIT_OF_DWORD : BOOL
  VAR_INPUT
    IN : DWORD;
    N : INT;
  END_VAR

  BIT_OF_DWORD := (SHR(in,N) AND 16#00000001) > 0;
  (* from OSCAT library; www.oscat.de  *)
END_FUNCTION

FUNCTION_BLOCK FILL_Block
	VAR_INPUT
		C :	BYTE;
		L :	INT;
	END_VAR

	VAR_OUTPUT
		FILL :	STRING;
	END_VAR

	VAR
		N :	BYTE;
		I :	INT;
		sx :	STRING;
		CHR_TO_STRING :	CHR_TO_STRING_Block;
		FILL_tmp :	STRING;
	END_VAR

	CHR_TO_STRING(C:=c);
	Sx:=CHR_TO_STRING.CHR_TO_STRING;
	(* create string *)
	N := INT_TO_BYTE(LIMIT(0,L,80));
	(* create a string of characters to be connected to str *)
	FILL := '';
	FOR i := 1 TO 8 DO
		FILL_tmp := FILL;
		FILL := CONCAT(FILL_tmp,FILL);
		IF BIT_OF_DWORD(BYTE_TO_DWORD(N),7) THEN FILL := CONCAT(FILL,Sx); END_IF;
		N := SHL(N,1);
	END_FOR;
END_FUNCTION_BLOCK

PROGRAM program0
  VAR
	C :	BYTE;
	L :	INT;

	FILL :	STRING;

	func_block : FILL_Block;
  END_VAR
	func_block.C  :=C ;
	func_block.L  :=L ;
	func_block();
	FILL := func_block.FILL;
END_PROGRAM

CONFIGURATION Config0
  RESOURCE Res0 ON PLC
    TASK task0(INTERVAL := T#20ms,PRIORITY := 0);
    PROGRAM instance0 WITH task0 : program0;
  END_RESOURCE
END_CONFIGURATION

(* ---- 428-STACK_32.ST ---- *)
TYPE
  	oscat_ardw_0_31             : ARRAY [0..31]   OF DWORD;
END_TYPE

FUNCTION_BLOCK STACK_32_Block

	VAR_INPUT
		DIN :	DWORD;
		E :	BOOL := TRUE;
		RD :	BOOL;
		WD :	BOOL;
		RST :	BOOL;
	END_VAR

	VAR_OUTPUT
		DOUT :	DWORD;
		EMPTY :	BOOL := TRUE;
		FULL :	BOOL;
	END_VAR

	VAR
		pt :	INT;
		stack :	oscat_ardw_0_31;
	END_VAR

	IF RST THEN
		pt := 0;
		EMPTY := TRUE;
		FULL := FALSE;
		Dout := DWORD#0;
	ELSIF E THEN
		IF NOT EMPTY AND RD THEN
			(* read one element *)
			pt := pt - 1;
			Dout := stack[pt];
			EMPTY := pt = 0;
			FULL := FALSE;
		END_IF;
		IF NOT FULL AND WD THEN
			(* write one element *)
			stack[pt] := Din;
			pt := pt + 1;
			FULL := pt > 31;
			EMPTY := FALSE;
		END_IF;
	END_IF;

END_FUNCTION_BLOCK

PROGRAM program0
	VAR
		DIN :	DWORD;
		E :	BOOL := TRUE;
		RD :	BOOL;
		WD :	BOOL;
		RST :	BOOL;
		DOUT :	DWORD;
		EMPTY :	BOOL := TRUE;
		FULL :	BOOL;
		func_block : STACK_32_Block;
	END_VAR
		func_block.DIN  := DIN;
		func_block.E  := E;
		func_block.RD  := RD;
		func_block.WD  := WD;
		func_block.RST  := RST;
		func_block();
		DOUT := func_block.DOUT;
		EMPTY := func_block.EMPTY;
		FULL := func_block.FULL;

END_PROGRAM

CONFIGURATION Config0

	RESOURCE Res0 ON PLC
		TASK task0(INTERVAL := T#20ms,PRIORITY := 0);
		PROGRAM instance0 WITH task0 : program0;
	END_RESOURCE

END_CONFIGURATION

(* ---- 429-BUFFER_INSERT_NW.ST ---- *)
TYPE
  oscat_NW_BUF_LONG  : ARRAY [0..4095] OF BYTE;
END_TYPE

FUNCTION_BLOCK _BUFFER_INSERT_NW
	VAR_INPUT
		STR :	STRING;
		POS :	INT;
	END_VAR

	VAR_IN_OUT
		PT :	oscat_NW_BUF_LONG;
	END_VAR

	VAR_INPUT
		SIZE :	UINT;
	END_VAR

	VAR_OUTPUT
		_BUFFER_INSERT :	INT;
	END_VAR

	VAR
		end :	INT;
		lx :	INT;
		i :	INT;
		i2 :	INT;
		_STRING_TO_BUFFER :	_STRING_TO_BUFFER;
	END_VAR

	i := UINT_TO_INT(size) - 1;
	pos := LIMIT_INT(0,pos,i);
	lx := LEN(str);
	end := pos + lx;
	(* first move the upper part of the buffer to make space for the string *)
	i2 := i - lx;
	WHILE i >= end DO
	pt[i] := pt[i2];
	i  := i  - 1;
	i2 := i2 - 1;
	END_WHILE;

	_STRING_TO_BUFFER(str:=str, pos:=pos, size:=size, pt:=pt);
	_BUFFER_INSERT := _STRING_TO_BUFFER._STRING_TO_BUFFER;
	pt := _STRING_TO_BUFFER.pt;
END_FUNCTION_BLOCK

PROGRAM program0
  VAR
	STR :	STRING;
	POS :	INT;

	PT :	oscat_NW_BUF_LONG;

	SIZE :	UINT;

	_BUFFER_INSERT :	INT;
	func_block : _BUFFER_INSERT_NW;
  END_VAR
	func_block.STR  :=STR ;
	func_block.POS  :=POS ;
	func_block.SIZE  :=SIZE ;
	func_block.PT  :=PT ;
	func_block();
	PT := func_block.PT;
	_BUFFER_INSERT := func_block._BUFFER_INSERT;
END_PROGRAM

CONFIGURATION Config0
  RESOURCE Res0 ON PLC
    TASK task0(INTERVAL := T#20ms,PRIORITY := 0);
    PROGRAM instance0 WITH task0 : program0;
  END_RESOURCE
END_CONFIGURATION

(* ---- 430-_BUFFER_UPPERCASE_NW.ST ---- *)
TYPE
  oscat_NW_BUF_LONG  : ARRAY [0..4095] OF BYTE;
END_TYPE

FUNCTION SETUP_EXTENDED_ASCII:BOOL
	VAR_INPUT
		X :	BOOL;
	END_VAR

	SETUP_EXTENDED_ASCII := X OR TRUE;
END_FUNCTION

FUNCTION TO_UPPER:BYTE

	VAR_INPUT
		IN :	BYTE;
	END_VAR

	IF in > BYTE#96 AND in < BYTE#123 THEN
	TO_UPPER := in AND BYTE#16#DF;
	ELSIF in > BYTE#223 AND in <> BYTE#247 AND in <> BYTE#255 AND SETUP_EXTENDED_ASCII(FALSE) THEN
	TO_UPPER := in AND BYTE#16#DF;
	ELSE
	TO_UPPER := in;
	END_IF;

END_FUNCTION

FUNCTION_BLOCK _BUFFER_UPPERCASE_NW
	VAR_INPUT
		SIZE :	UINT;
	END_VAR

	VAR_OUTPUT
		_BUFFER_UPPERCASE :	BOOL;
	END_VAR

	VAR_IN_OUT
		PT :	oscat_NW_BUF_LONG;
	END_VAR

	VAR
		pos :	INT;
		size2 :	INT;
	END_VAR

	pos := 0;
	size2 := UINT_TO_INT(SIZE);

	WHILE pos < size2 DO
		PT[pos] := TO_UPPER(PT[pos]);
		pos := pos + 1;
	END_WHILE;

	_BUFFER_UPPERCASE := TRUE;

END_FUNCTION_BLOCK

PROGRAM program0
  VAR
	SIZE :	UINT;

	_BUFFER_UPPERCASE :	BOOL;

	PT :	oscat_NW_BUF_LONG;

	func_block : _BUFFER_UPPERCASE_NW;
  END_VAR
	func_block.SIZE  :=SIZE ;
	func_block.PT  :=PT ;
	func_block();
	PT := func_block.PT;
	_BUFFER_UPPERCASE := func_block._BUFFER_UPPERCASE;
END_PROGRAM

CONFIGURATION Config0
  RESOURCE Res0 ON PLC
    TASK task0(INTERVAL := T#20ms,PRIORITY := 0);
    PROGRAM instance0 WITH task0 : program0;
  END_RESOURCE
END_CONFIGURATION

(* ---- 431-SCHEDULER_2.ST ---- *)
FUNCTION_BLOCK SCHEDULER_2_Block

	VAR_INPUT
		E0 :	BOOL;
		E1 :	BOOL;
		E2 :	BOOL;
		E3 :	BOOL;
		C0 :	UINT;
		C1 :	UINT;
		C2 :	UINT;
		C3 :	UINT;
		O0 :	UINT;
		O1 :	UINT;
		O2 :	UINT;
		O3 :	UINT;
	END_VAR

	VAR_OUTPUT
		Q0 :	BOOL;
		Q1 :	BOOL;
		Q2 :	BOOL;
		Q3 :	BOOL;
	END_VAR

	VAR
		sx :	UINT;
	END_VAR

	Q0 := E0 AND (sx MOD C0 - O0 = UINT#0);
	Q1 := E1 AND (sx MOD C1 - O1 = UINT#0);
	Q2 := E2 AND (sx MOD C2 - O2 = UINT#0);
	Q3 := E3 AND (sx MOD C3 - O3 = UINT#0);

	sx := sx + UINT#1;

END_FUNCTION_BLOCK

PROGRAM program0

	VAR
		E0 :	BOOL;
		E1 :	BOOL;
		E2 :	BOOL;
		E3 :	BOOL;
		C0 :	UINT;
		C1 :	UINT;
		C2 :	UINT;
		C3 :	UINT;
		O0 :	UINT;
		O1 :	UINT;
		O2 :	UINT;
		O3 :	UINT;
		Q0 :	BOOL;
		Q1 :	BOOL;
		Q2 :	BOOL;
		Q3 :	BOOL;
		func_block : SCHEDULER_2_Block;
  	END_VAR
	func_block.E0  :=	E0;
	func_block.E1  :=	E1;
	func_block.E2  :=	E2;
	func_block.E3  :=	E3;
	func_block.C0  :=	C0;
	func_block.C1  :=	C1;
	func_block.C2  :=	C2;
	func_block.C3  :=	C3;
	func_block.O0  :=	O0;
	func_block.O1  :=	O1;
	func_block.O2  :=	O2;
	func_block.O3  :=	O3;
	func_block();
	Q0 := func_block.Q0;
	Q1 := func_block.Q1;
	Q2 := func_block.Q2;
	Q3 := func_block.Q3;

END_PROGRAM

CONFIGURATION Config0

	RESOURCE Res0 ON PLC
		TASK task0(INTERVAL := T#20ms,PRIORITY := 0);
		PROGRAM instance0 WITH task0 : program0;
	END_RESOURCE

END_CONFIGURATION

(* ---- 432-BYTE_TO_BITS.ST ---- *)
FUNCTION BIT_OF_DWORD : BOOL
  VAR_INPUT
    IN : DWORD;
    N : INT;
  END_VAR

  BIT_OF_DWORD := (SHR(in,N) AND 16#00000001) > 0;
END_FUNCTION

FUNCTION_BLOCK BYTE_TO_BITS
	VAR_INPUT
		IN :	BYTE;
	END_VAR

	VAR_OUTPUT
		B0 :	BOOL;
		B1 :	BOOL;
		B2 :	BOOL;
		B3 :	BOOL;
		B4 :	BOOL;
		B5 :	BOOL;
		B6 :	BOOL;
		B7 :	BOOL;
	END_VAR

	B0 := BIT_OF_DWORD(BYTE_TO_DWORD(IN),0); (* IN.X0 *)
	B1 := BIT_OF_DWORD(BYTE_TO_DWORD(IN),1); (* IN.X1 *)
	B2 := BIT_OF_DWORD(BYTE_TO_DWORD(IN),2); (* IN.X2 *)
	B3 := BIT_OF_DWORD(BYTE_TO_DWORD(IN),3); (* IN.X3 *)
	B4 := BIT_OF_DWORD(BYTE_TO_DWORD(IN),4); (* IN.X4 *)
	B5 := BIT_OF_DWORD(BYTE_TO_DWORD(IN),5); (* IN.X5 *)
	B6 := BIT_OF_DWORD(BYTE_TO_DWORD(IN),6); (* IN.X6 *)
	B7 := BIT_OF_DWORD(BYTE_TO_DWORD(IN),7); (* IN.X7 *)
END_FUNCTION_BLOCK

PROGRAM program0
  VAR
	LocalVar0  : BYTE;
	B0 :	BOOL;
	B1 :	BOOL;
	B2 :	BOOL;
	B3 :	BOOL;
	B4 :	BOOL;
	B5 :	BOOL;
	B6 :	BOOL;
	B7 :	BOOL;
	func_block: BYTE_TO_BITS;
  END_VAR

	func_block.IN  := LocalVar0;
	func_block();
	B0 := func_block.B0;
	B1 := func_block.B1;
	B2 := func_block.B2;
	B3 := func_block.B3;
	B4 := func_block.B4;
	B5 := func_block.B5;
	B6 := func_block.B6;
	B7 := func_block.B7;

END_PROGRAM

CONFIGURATION Config0
  RESOURCE Res0 ON PLC
    TASK task0(INTERVAL := T#20ms,PRIORITY := 0);
    PROGRAM instance0 WITH task0 : program0;
  END_RESOURCE
END_CONFIGURATION

(* ---- 433-LOG_MSG.ST ---- *)
FUNCTION_BLOCK LOG_MSG

	VAR_EXTERNAL
		LOG_CL :	us_LOG_CONTROL;
	END_VAR

	VAR
		FB_PRINT_SF :	PRINT_SF;
		idx :	INT;
	END_VAR

	IF DWORD_TO_BYTE(SHL(LOG_CL.NEW_MSG_OPTION,16)) > LOG_CL.LEVEL THEN RETURN; END_IF;
	LOG_CL.SIZE := 400;

	FB_PRINT_SF.PRINTF_DATA := LOG_CL.PRINTF;
	FB_PRINT_SF.STR 		:= LOG_CL.NEW_MSG;
	FB_PRINT_SF();
	LOG_CL.NEW_MSG	:= FB_PRINT_SF.STR;
	LOG_CL.PRINTF	:= FB_PRINT_SF.PRINTF_DATA;

	IF LOG_CL.RESET THEN
		LOG_CL.RESET := FALSE;
		LOG_CL.RING_MODE := FALSE;
		LOG_CL.IDX := 0;
		LOG_CL.UPDATE_COUNT := LOG_CL.UPDATE_COUNT + UINT#1;
	END_IF;

	IF LOG_CL.SIZE > 0 THEN
		IF LEN(LOG_CL.NEW_MSG) > 0 THEN
			IF (LOG_CL.IDX >= LOG_CL.SIZE) THEN
				LOG_CL.RING_MODE := TRUE;
				LOG_CL.IDX := 0;
			END_IF;

			LOG_CL.UPDATE_COUNT := LOG_CL.UPDATE_COUNT + UINT#1;
			LOG_CL.IDX := LOG_CL.IDX + INT#1;
			idx := LOG_CL.IDX;
			LOG_CL.MSG[idx] := LOG_CL.NEW_MSG;
			LOG_CL.MSG_OPTION[idx] := LOG_CL.NEW_MSG_OPTION;
			LOG_CL.NEW_MSG := '';
		END_IF;
	END_IF;

END_FUNCTION_BLOCK

PROGRAM program0
	VAR
		STR :	oscat_STRING80;
		LOG_MSG_R :	DWORD;
		func_block : LOG_MSG;
	END_VAR

	func_block.STR := STR;
	func_block();
	LOG_MSG_R  := func_block.LOG_MSG;
END_PROGRAM

CONFIGURATION Config0
  	RESOURCE Res0 ON PLC
    	TASK task0(INTERVAL := T#20ms,PRIORITY := 0);
    	PROGRAM instance0 WITH task0 : program0;
  	END_RESOURCE
END_CONFIGURATION

(* ---- 434-ARRAY_SDV.ST ---- *)
TYPE
	oscat_pt_ARRAY: ARRAY [1..100] OF REAL;
END_TYPE

FUNCTION_BLOCK ARRAY_VAR_Block
	VAR_IN_OUT
		PT :	oscat_pt_ARRAY;
	END_VAR

	VAR_INPUT
		SIZE :	UINT;
	END_VAR

	VAR_OUTPUT
		ARRAY_VAR :	REAL;
	END_VAR

	VAR
		i :	INT;
		stop :	INT;
		avg :	REAL;
	END_VAR

	stop :=LIMIT_INT(1,UINT_TO_INT(size),1000);
	avg := pt[1];
	FOR i := 2 TO stop DO
		avg := avg + pt[i];
	END_FOR;
	avg := avg / INT_TO_REAL(stop);

	array_var := EXPT(pt[1] - avg, 2.0);
	FOR i := 2 TO stop DO
		array_var := array_var + EXPT(pt[i] - avg, 2.0);
	END_FOR;
	array_var := array_var / INT_TO_REAL(stop-1);

END_FUNCTION_BLOCK

FUNCTION_BLOCK ARRAY_SDV_Block
	VAR_IN_OUT
		PT :	oscat_pt_ARRAY;
	END_VAR

	VAR_INPUT
		SIZE :	UINT;
	END_VAR

	VAR_OUTPUT
		ARRAY_SDV :	REAL;
	END_VAR

	VAR
		FB_array_var :	array_var_block;
	END_VAR

	FB_array_var.pt   := pt;
	FB_array_var.size := size;
	FB_array_var();
	pt := FB_array_var.pt;

	array_sdv := SQRT(FB_array_var.array_var);
END_FUNCTION_BLOCK

PROGRAM program0
  VAR
    LocalVar0 : oscat_pt_ARRAY;
    LocalVar1 : UINT;
	LocalOUT  : REAL;
	func_block : ARRAY_SDV_Block;
  END_VAR
	func_block.pt := LocalVar0;
	func_block.size := LocalVar1;
	func_block();
	LocalOUT := func_block.ARRAY_SDV;

END_PROGRAM

CONFIGURATION Config0
  RESOURCE Res0 ON PLC
    TASK task0(INTERVAL := T#20ms,PRIORITY := 0);
    PROGRAM instance0 WITH task0 : program0;
  END_RESOURCE
END_CONFIGURATION

(* ---- 435-FIFO_16.ST ---- *)
TYPE
	oscat_ardw_0_15             : ARRAY [0..15]   OF DWORD;
END_TYPE

FUNCTION INC1:INT

	VAR_INPUT
		X :	INT;
		N :	INT;
	END_VAR

	IF X >= N - 1 THEN
		INC1 := 0;
	ELSE
		INC1 := X + 1;
	END_IF;
END_FUNCTION

FUNCTION_BLOCK FIFO_16
	VAR_INPUT
		DIN :	DWORD;
		E :	BOOL := TRUE;
		RD :	BOOL;
		WD :	BOOL;
		RST :	BOOL;
	END_VAR

	VAR_OUTPUT
		DOUT :	DWORD;
		EMPTY :	BOOL := TRUE;
		FULL :	BOOL;
	END_VAR

	VAR
		fifo :	oscat_ardw_0_15;
		pr :	INT;
		pw :	INT;
	END_VAR

	IF RST THEN
		pw := pr;
		FULL := FALSE;
		EMPTY := TRUE;
		Dout := DWORD#0;
	ELSIF E THEN
		IF NOT EMPTY AND RD THEN
			Dout := fifo[pr];
			pr := INC1(pr,16);
			EMPTY := pr = pw;
			FULL := FALSE;
		END_IF;
		IF NOT FULL AND WD THEN
			fifo[pw] := Din;
			pw := INC1(pw,16);
			FULL := pw = pr;
			EMPTY := FALSE;
		END_IF;
	END_IF;
END_FUNCTION_BLOCK

PROGRAM program0
  VAR
	DIN :	DWORD;
	E   :	BOOL;
	RD  :	BOOL;
	WD  :	BOOL;
	RST :	BOOL;

	DOUT  :	DWORD;
	EMPTY :	BOOL;
	FULL  :	BOOL;

	func_block : FIFO_16;
  END_VAR
	func_block.DIN :=DIN;
	func_block.E   :=E  ;
	func_block.RD  :=RD ;
	func_block.WD  :=WD ;
	func_block.RST :=RST;
	func_block();
	DOUT := func_block.DOUT ;
	EMPTY:= func_block.EMPTY;
	FULL := func_block.FULL ;
END_PROGRAM

CONFIGURATION Config0
  RESOURCE Res0 ON PLC
    TASK task0(INTERVAL := T#20ms,PRIORITY := 0);
    PROGRAM instance0 WITH task0 : program0;
  END_RESOURCE
END_CONFIGURATION

(* ---- 437-CCOS.ST ---- *)
TYPE oscat_complex :
  STRUCT
	re : REAL;
	im : REAL;
  END_STRUCT;
END_TYPE

FUNCTION COSH:REAL
	VAR_INPUT
		X :	REAL;
	END_VAR

	VAR
		t :	REAL;
	END_VAR

	T := EXP(X);
	COSH := (1.0 / T + T) * 0.5;
END_FUNCTION

FUNCTION SINH:REAL
	VAR_INPUT
		X :	REAL;
	END_VAR

	IF ABS(x) < 2.0E-3 THEN
		SINH := X;
	ELSE
		SINH := (EXP(x) - EXP(-x)) * 0.5;
	END_IF;
END_FUNCTION

FUNCTION_BLOCK CCOSH_Block
	VAR_INPUT
		X :	oscat_complex;
	END_VAR

	VAR_OUTPUT
		CCOSH :	oscat_complex;
	END_VAR

	CCOSH.re := cosH(x.re) * COS(x.im);
	CCOSH.im := sinH(x.re) * SIN(x.im);
END_FUNCTION_BLOCK

FUNCTION_BLOCK CSET_Block
	VAR_INPUT
		RE :	REAL;
		IM :	REAL;
	END_VAR

	VAR_OUTPUT
		CSET :	oscat_complex;
	END_VAR

	CSET.re := RE;
	CSET.im := IM;
END_FUNCTION_BLOCK

FUNCTION_BLOCK CCOS_Block
	VAR_INPUT
		X :	oscat_complex;
	END_VAR

	VAR_OUTPUT
		CCOS :	oscat_complex;
	END_VAR

	VAR
		CSET :	CSET_Block;
		CCOSH :	CCOSH_Block;
	END_VAR

	CSET(RE:= -X.im,IM:=X.re);
	CCOSH(X:=CSET.CSET);
	CCOS := CCOSH.CCOSH;

END_FUNCTION_BLOCK

PROGRAM program0
  VAR
    LocalVar0 : oscat_complex;
	LocalOUT  : oscat_complex;
	func_block : CCOS_Block;
  END_VAR
	func_block.X  := LocalVar0;
	func_block();
	LocalOUT := func_block.CCOS;
END_PROGRAM

CONFIGURATION Config0
  RESOURCE Res0 ON PLC
    TASK task0(INTERVAL := T#20ms,PRIORITY := 0);
    PROGRAM instance0 WITH task0 : program0;
  END_RESOURCE
END_CONFIGURATION

(* ---- 438-FIFO_32.ST ---- *)
TYPE
	oscat_ardw_0_31             : ARRAY [0..31]   OF DWORD;
END_TYPE

FUNCTION INC1:INT

	VAR_INPUT
		X :	INT;
		N :	INT;
	END_VAR

	IF X >= N - 1 THEN
		INC1 := 0;
	ELSE
		INC1 := X + 1;
	END_IF;
END_FUNCTION

FUNCTION_BLOCK FIFO_32

	VAR_INPUT
		DIN :	DWORD;
		E :	BOOL := TRUE;
		RD :	BOOL;
		WD :	BOOL;
		RST :	BOOL;
	END_VAR

	VAR_OUTPUT
		DOUT :	DWORD;
		EMPTY :	BOOL := TRUE;
		FULL :	BOOL;
	END_VAR

	VAR
		fifo :	oscat_ardw_0_31;
		pr :	INT;
		pw :	INT;
	END_VAR

	IF RST THEN
		pw := pr;
		FULL := FALSE;
		EMPTY := TRUE;
		Dout := DWORD#0;
	ELSIF E THEN
		IF NOT EMPTY AND RD THEN
			Dout := fifo[pr];
			pr := INC1(pr,32);
			EMPTY := pr = pw;
			FULL := FALSE;
		END_IF;
		IF NOT FULL AND WD THEN
			fifo[pw] := Din;
			pw := INC1(pw,32);
			FULL := pw = pr;
			EMPTY := FALSE;
		END_IF;
	END_IF;

END_FUNCTION_BLOCK

PROGRAM program0
  VAR
	DIN :	DWORD;
	E   :	BOOL;
	RD  :	BOOL;
	WD  :	BOOL;
	RST :	BOOL;

	DOUT  :	DWORD;
	EMPTY :	BOOL;
	FULL  :	BOOL;

	func_block : FIFO_32;
  END_VAR
	func_block.DIN :=DIN;
	func_block.E   :=E  ;
	func_block.RD  :=RD ;
	func_block.WD  :=WD ;
	func_block.RST :=RST;
	func_block();
	DOUT := func_block.DOUT ;
	EMPTY:= func_block.EMPTY;
	FULL := func_block.FULL ;
END_PROGRAM

CONFIGURATION Config0
  RESOURCE Res0 ON PLC
    TASK task0(INTERVAL := T#20ms,PRIORITY := 0);
    PROGRAM instance0 WITH task0 : program0;
  END_RESOURCE
END_CONFIGURATION

(* ---- 439-ALARM_2.ST ---- *)
FUNCTION_BLOCK ALARM_2
	VAR_INPUT
		X :	REAL;
		LO_1 :	REAL;
		HI_1 :	REAL;
		LO_2 :	REAL;
		HI_2 :	REAL;
		HYS :	REAL;
	END_VAR

	VAR_OUTPUT
		Q1_LO :	BOOL;
		Q1_HI :	BOOL;
		Q2_LO :	BOOL;
		Q2_HI :	BOOL;
	END_VAR

	VAR
		tmp :	REAL;
	END_VAR

	tmp := X - Hys * 0.5;
	IF tmp > LO_1 THEN Q1_LO := FALSE; END_IF;
	IF tmp > LO_2 THEN Q2_LO := FALSE; END_IF;
	IF tmp > HI_1 THEN Q1_HI := TRUE; END_IF;
	IF tmp > HI_2 THEN Q2_HI := TRUE; END_IF;
	tmp := tmp + hys;
	IF tmp < LO_1 THEN Q1_LO := TRUE; END_IF;
	IF tmp < LO_2 THEN Q2_LO := TRUE; END_IF;
	IF tmp < HI_1 THEN Q1_HI := FALSE; END_IF;
	IF tmp < HI_2 THEN Q2_HI := FALSE; END_IF;

END_FUNCTION_BLOCK

PROGRAM program0
	VAR
	    LocalVar0 : REAL;
		LocalVar1 : REAL;
		LocalVar2 : REAL;
		LocalVar3 : REAL;
		LocalVar4 : REAL;
		LocalVar5 : REAL;
		LocalOUT1  : BOOL;
		LocalOUT2  : BOOL;
		LocalOUT3  : BOOL;
		LocalOUT4  : BOOL;
		func_block : ALARM_2;
  	END_VAR
	func_block.X := LocalVar0;
	func_block.LO_1 := LocalVar1;
	func_block.HI_1 := LocalVar2;
	func_block.LO_2 := LocalVar3;
	func_block.HI_2 := LocalVar4;
	func_block.HYS := LocalVar5;
	func_block();
	LocalOUT1 := func_block.Q1_LO;
	LocalOUT2 := func_block.Q1_HI;
	LocalOUT3 := func_block.Q2_LO;
	LocalOUT4 := func_block.Q2_HI;
END_PROGRAM

CONFIGURATION Config0
  	RESOURCE Res0 ON PLC
    	TASK task0(INTERVAL := T#20ms,PRIORITY := 0);
    	PROGRAM instance0 WITH task0 : program0;
  	END_RESOURCE
END_CONFIGURATION

(* ---- 440-DRIVER_4C.ST ---- *)
TYPE
  oscat_DRIVER_4C 			  : ARRAY [1..7] 	OF BYTE;
END_TYPE
FUNCTION_BLOCK DRIVER_4C

	VAR_INPUT
		IN :	BOOL;
		RST :	BOOL;
		TIMEOUT :	TIME;
		SX :	oscat_DRIVER_4C;
	END_VAR

	VAR_OUTPUT
		SN :	INT;
		Q0 :	BOOL;
		Q1 :	BOOL;
		Q2 :	BOOL;
		Q3 :	BOOL;
	END_VAR

	VAR
		off :	TON;
		edge :	BOOL;
	END_VAR

	IF RST OR off.Q THEN
		SN := 0;
	ELSIF IN AND NOT edge THEN
		SN := SN + 1;
		IF SN > 7 OR SX[SN] = BYTE#0 THEN SN := 0; END_IF;
	END_IF;
	edge := in;
	IF SN > 0 THEN
		Q0 := (SX[SN] AND BYTE#1) > BYTE#0;
		Q1 := (SX[SN] AND BYTE#2) > BYTE#0;
		Q2 := (SX[SN] AND BYTE#4) > BYTE#0;
		Q3 := (SX[SN] AND BYTE#8) > BYTE#0;
	ELSE
		Q0 := FALSE;
		Q1 := FALSE;
		Q2 := FALSE;
		Q3 := FALSE;
	END_IF;

	IF timeout > t#0s THEN off(in := SN > 0, PT := Timeout); END_IF;

END_FUNCTION_BLOCK

PROGRAM program0
  VAR
	IN      :	BOOL;
	RST     :	BOOL;
	TIMEOUT :	TIME;
	SX      :	oscat_DRIVER_4C;

	SN :	INT;
	Q0 :	BOOL;
	Q1 :	BOOL;
	Q2 :	BOOL;
	Q3 :	BOOL;

	func_block : DRIVER_4C;
  END_VAR
	func_block.IN       :=IN      ;
	func_block.RST      :=RST     ;
	func_block.TIMEOUT  :=TIMEOUT ;
	func_block.SX       :=SX      ;
	func_block();
	SN := func_block.SN;
	Q0 := func_block.Q0;
	Q1 := func_block.Q1;
	Q2 := func_block.Q2;
	Q3 := func_block.Q3;
END_PROGRAM

CONFIGURATION Config0
  RESOURCE Res0 ON PLC
    TASK task0(INTERVAL := T#20ms,PRIORITY := 0);
    PROGRAM instance0 WITH task0 : program0;
  END_RESOURCE
END_CONFIGURATION

(* ---- 441-COUNT_DR.ST ---- *)
FUNCTION_BLOCK COUNT_DR
	VAR_INPUT
		SET :	BOOL;
		IN :	DWORD;
		UP :	BOOL;
		DN :	BOOL;
		STEPP :	DWORD := DWORD#1;
		MX :	DWORD := DWORD#16#FFFF_FFFF;
		RST :	BOOL;
	END_VAR

	VAR_OUTPUT
		CNT :	DWORD;
	END_VAR

	VAR
		CNT2 :	UDINT;
		STEPP2 :	UDINT;
		MX2 :	UDINT;
		last_up :	BOOL;
		last_dn :	BOOL;
	END_VAR

	STEPP2 := DWORD_TO_UDINT(STEPP);
	MX2   := DWORD_TO_UDINT(MX);
	CNT2  := DWORD_TO_UDINT(CNT);

	IF rst THEN
		CNT2 := UDINT#0;
	ELSIF set THEN
		CNT2 := LIMIT(UDINT#0,DWORD_TO_UDINT(in),mx2);
	ELSIF up AND NOT last_up THEN
		IF STEPP2 > MX2 - CNT2 THEN
			CNT2 := CNT2 - MX2 + STEPP2 - UDINT#1;
		ELSE
			CNT2 := CNT2 + STEPP2;
		END_IF;
	ELSIF dn AND NOT last_dn THEN
		IF STEPP2 > CNT2 THEN
			CNT2 := CNT2 - STEPP2 + MX2 + UDINT#1;
		ELSE
			CNT2 := CNT2 - STEPP2;
		END_IF;
	END_IF;
	last_up := up;
	last_dn := dn;
	CNT := UDINT_TO_DWORD(CNT2);
END_FUNCTION_BLOCK

PROGRAM program0
  VAR
	SET :	BOOL;
	IN :	DWORD;
	UP :	BOOL;
	DN :	BOOL;
	STEPP :	DWORD;
	MX :	DWORD;
	RST :	BOOL;

	CNT :	DWORD;
	func_block : COUNT_DR;
  END_VAR
	func_block.SET  :=SET  ;
	func_block.IN   :=IN   ;
	func_block.UP   :=UP   ;
	func_block.DN   :=DN   ;
	func_block.STEPP :=STEPP ;
	func_block.MX   :=MX   ;
	func_block.RST  :=RST  ;

	func_block();
	CNT := func_block.CNT;
END_PROGRAM

CONFIGURATION Config0
  RESOURCE Res0 ON PLC
    TASK task0(INTERVAL := T#20ms,PRIORITY := 0);
    PROGRAM instance0 WITH task0 : program0;
  END_RESOURCE
END_CONFIGURATION

(* ---- 442-BUFFER_SEARCH.ST ---- *)
TYPE
	oscat_arb_0_249 			  : ARRAY [0..249] 	OF BYTE;
END_TYPE

FUNCTION_BLOCK BUFFER_SEARCH_Block
	VAR_INPUT
		SIZE :	UINT;
		STR :	STRING;
		POS :	INT;
		IGN :	BOOL;
	END_VAR

	VAR_IN_OUT
		PT :	oscat_arb_0_249;
	END_VAR

	VAR_OUTPUT
		BUFFER_SEARCH :	INT;
	END_VAR

	VAR
		i :	INT;
		end :	INT;
		k :	INT;
		k2 :	INT;
		lx :	INT;
		char :	BYTE;
		chx :	BYTE;
	END_VAR

	lx := LEN(str);
	IF pos >= 0 AND lx > 0 THEN
		end := UINT_TO_INT(size) - lx;
		lx := lx - 1;
		FOR i := pos TO end DO
			FOR k := 0 TO lx DO
				char := INT_TO_BYTE(GET_CHAR(str,k + 1));
				k2 := i + k;
				IF IGN THEN
					chx := TO_UPPER(pt[k2]);
				ELSE
					chx := pt[k2];
				END_IF;
				IF char <> chx THEN EXIT; END_IF;
			END_FOR;
			IF k > lx THEN
				BUFFER_SEARCH := i;
				RETURN;
			END_IF;
		END_FOR;
	END_IF;
	BUFFER_SEARCH := -1;
END_FUNCTION_BLOCK

PROGRAM program0
  VAR
    LocalVar0 : UINT;
    LocalVar1 : STRING;
	LocalVar2 : INT;
	LocalVar3 : BOOL;
	LocalVar4 : oscat_arb_0_249;
	LocalOUT  : INT;
	func_block : BUFFER_COMP_Block;
  END_VAR
	func_block.SIZE  := LocalVar0;
	func_block.STR  := LocalVar1;
	func_block.POS   := LocalVar2;
	func_block.IGN  := LocalVar3;
	func_block.PT := LocalVar4;
	func_block();
	LocalOUT := func_block.BUFFER_COMP;
	LocalVar4 := func_block.PT;

END_PROGRAM

CONFIGURATION Config0
  RESOURCE Res0 ON PLC
    TASK task0(INTERVAL := T#20ms,PRIORITY := 0);
    PROGRAM instance0 WITH task0 : program0;
  END_RESOURCE
END_CONFIGURATION

(* ---- 445-COUNT_BR.ST ---- *)
FUNCTION _BYTE_TO_INT:INT
	VAR_INPUT
		IN :	BYTE;
	END_VAR

	_BYTE_TO_INT := USINT_TO_INT(BYTE_TO_USINT(IN));

END_FUNCTION

FUNCTION INC:INT
	VAR_INPUT
		X :	INT;
		D :	INT;
		M :	INT;
	END_VAR

	inc := (X + D + M + 1) MOD (M + 1);
END_FUNCTION

FUNCTION_BLOCK COUNT_BR
	VAR_INPUT
		SET :	BOOL;
		IN :	BYTE;
		UP :	BOOL;
		DN :	BOOL;
		STEPP :	BYTE := BYTE#1;
		MX :	BYTE := BYTE#255;
		RST :	BOOL;
	END_VAR
	VAR_OUTPUT
		CNT :	BYTE;
	END_VAR

	VAR
		last_up :	BOOL;
		last_dn :	BOOL;
	END_VAR

	IF rst THEN
		cnt := BYTE#0;
	ELSIF set THEN
		cnt := INT_TO_BYTE(LIMIT(0,_BYTE_TO_INT(in),_BYTE_TO_INT(mx)));
	ELSIF up AND NOT last_up THEN
		cnt := INT_TO_BYTE(inc(_BYTE_TO_INT(cnt),_BYTE_TO_INT(stepP),_BYTE_TO_INT(mx)));
	ELSIF dn AND NOT last_dn THEN
		cnt := INT_TO_BYTE(inc(_BYTE_TO_INT(cnt),_BYTE_TO_INT(stepP) * -1,_BYTE_TO_INT(mx)));
	END_IF;
	last_up := up;
	last_dn := dn;
END_FUNCTION_BLOCK

PROGRAM program0
  VAR
	SET :	BOOL;
	IN :	BYTE;
	UP :	BOOL;
	DN :	BOOL;
	STEPP:	BYTE;
	MX :	BYTE;
	RST :	BOOL;

	CNT :	BYTE;
	func_block : COUNT_BR;
  END_VAR
	func_block.SET  :=SET  ;
	func_block.IN   :=IN   ;
	func_block.UP   :=UP   ;
	func_block.DN   :=DN   ;
	func_block.STEPP :=STEPP ;
	func_block.MX   :=MX   ;
	func_block.RST  :=RST  ;

	func_block();
	CNT := func_block.CNT;
END_PROGRAM

CONFIGURATION Config0
  RESOURCE Res0 ON PLC
    TASK task0(INTERVAL := T#20ms,PRIORITY := 0);
    PROGRAM instance0 WITH task0 : program0;
  END_RESOURCE
END_CONFIGURATION

(* ---- 446-RC4_CRYPT_STREAM.ST ---- *)
FUNCTION_BLOCK RC4_CRYPT_STREAM

	VAR_IN_OUT
		MODE :	INT;
		KEY :	oscat_STRING40;
		BUF :	oscat_aB0_63;
		SIZE :	UDINT;
	END_VAR

	VAR_OUTPUT
		POS :	UDINT;
	END_VAR

	VAR
		sbox :	oscat_aB0_255;
		skey :	oscat_aB0_255;
		a :	INT;
		b :	INT;
		c :	INT;
		d :	USINT;
		e :	USINT;
		end :	UDINT;
		v :	BYTE;
		v_tmp :	INT;
		CODE :	CODE;
	END_VAR

	CASE MODE OF

	1:
		b := LEN(KEY) - 1;
		IF b < 0 OR SIZE < UDINT#1 THEN
			MODE := 3;
			RETURN;
		END_IF;

		FOR a := 0 TO b DO
			CODE(STR:=KEY,POS:=a + 1);
			skey[a] := CODE.CODE;
			sbox[a] := INT_TO_BYTE(a);
		END_FOR;

		c := 0;
		FOR a := b + 1 TO 255 DO
			skey[a] := skey[c];
			sbox[a] := INT_TO_BYTE(a);
			c := c + 1;
			IF c > b THEN c := 0; END_IF;
		END_FOR;

		d := USINT#0;
		FOR a := 0 TO 255 DO
			d := d + BYTE_TO_USINT(sbox[a]) + BYTE_TO_USINT(skey[a]);
			v := sbox[a];
			sbox[a] := sbox[d];
			sbox[d] := v;
		END_FOR;

		POS := UDINT#0;
		end := SIZE;
		SIZE := MIN(UDINT#64,end);
		d := USINT#0;
		e := USINT#0;
		MODE := 2;

	2:

		b := UDINT_TO_INT(SIZE) - 1;
		FOR a := 0 TO b DO
			d := d + USINT#1;
			e := e + BYTE_TO_USINT(sbox[d]);
			v := sbox[d];
			sbox[d] := sbox[e];
			sbox[e] := v;
			v := USINT_TO_BYTE(BYTE_TO_USINT(sbox[d]) + BYTE_TO_USINT(sbox[e]));
			v_tmp := _BYTE_TO_INT(v);
			BUF[a] :=BUF[a] XOR sbox[v_tmp];
		END_FOR;

		POS := POS + SIZE;
		SIZE := MIN(UDINT#64,end - POS);

		IF SIZE = UDINT#0 THEN
			MODE := 3;
		END_IF;
	END_CASE;

END_FUNCTION_BLOCK

(* ---- 448-T_PLC_US.ST ---- *)
FUNCTION_BLOCK T_PLC_US_Block

	VAR_OUTPUT
		T_PLC_US :	UDINT;
	END_VAR

	VAR_EXTERNAL
		PLC_TICKS_PER_SEC :	INT;
		PLC_SYS_TICK_CNT :	DINT;
	END_VAR

	VAR
		debug :	BOOL;
		N :	INT;
		Offset :	UDINT;
		temp :	DWORD := DWORD#1;
		mode :	BOOL;
		faktor :	UDINT;
		init :	BOOL;
		v_plc_ticks_per_sec :	UDINT;
		base :	UDINT := UDINT#1000000;
	END_VAR

	IF init = FALSE THEN
		v_plc_ticks_per_sec := INT_TO_UDINT(PLC_TICKS_PER_SEC);
		IF v_plc_ticks_per_sec = UDINT#1024 THEN
			faktor := UDINT#1000;
			mode := FALSE;
		ELSIF v_plc_ticks_per_sec > UDINT#0 THEN
			IF v_plc_ticks_per_sec <= base THEN
				faktor := base / v_plc_ticks_per_sec;
				mode := FALSE;
			ELSE
				faktor := v_plc_ticks_per_sec / base;
				mode := TRUE;
			END_IF;
		ELSE
			faktor := UDINT#1;
		END_IF;
		init := TRUE;
	END_IF;

	IF mode THEN
		T_PLC_US := DINT_TO_UDINT(PLC_SYS_TICK_CNT) / faktor;
	ELSE
		T_PLC_US := DINT_TO_UDINT(PLC_SYS_TICK_CNT) * faktor;
	END_IF;

	IF debug THEN
		T_PLC_US := (DWORD_TO_UDINT(SHL(UDINT_TO_DWORD(T_PLC_US),N) OR SHL(temp,N)) - UDINT#1) + Offset;
	END_IF;

END_FUNCTION_BLOCK

PROGRAM program0

	VAR
		T_PLC_US  : UDINT;
		func_block : T_PLC_US_Block;
	END_VAR
		func_block();
		T_PLC_US := func_block.T_PLC_US;

END_PROGRAM

CONFIGURATION Config0

	VAR_GLOBAL
		PLC_TICKS_PER_SEC :	INT;
		PLC_SYS_TICK_CNT :	DINT;
	END_VAR

	RESOURCE Res0 ON PLC
		TASK task0(INTERVAL := T#20ms,PRIORITY := 0);
		PROGRAM instance0 WITH task0 : program0;
	END_RESOURCE

END_CONFIGURATION

(* ---- 449-REAL_TO_STRF.ST ---- *)
FUNCTION EXP10 : REAL

	VAR_INPUT
		x : REAL;
	END_VAR

	exp10 := EXP(X * 2.30258509299405);

END_FUNCTION

FUNCTION _REAL_TO_DINT:DINT
	VAR_INPUT
		X :	REAL;
	END_VAR

	IF REAL_TO_DINT(0.5) = DINT#1 THEN
		_REAL_TO_DINT := REAL_TO_DINT(x);
		RETURN;
	END_IF;

	IF X > 0.0 THEN
		_REAL_TO_DINT := REAL_TO_DINT(x+0.5);
	ELSIF X < 0.0 THEN
		_REAL_TO_DINT := REAL_TO_DINT(x-0.5);
	ELSE
		_REAL_TO_DINT := DINT#0;
	END_IF;
END_FUNCTION

FUNCTION_BLOCK REAL_TO_STRF_Block

	VAR_INPUT
		IN :	REAL;
		N :	INT;
		D :	STRING;
	END_VAR

	VAR_OUTPUT
		REAL_TO_STRF :	STRING;
	END_VAR

	VAR
		st_tmp : STRING;
		i :	INT;
	END_VAR

	N := LIMIT(0,N,7);
	REAL_TO_STRF := DINT_TO_STRING(_REAL_TO_DINT(ABS(in) * EXP10(INT_TO_REAL(N))));
	FOR i := LEN(REAL_TO_STRF) TO N DO
		st_tmp := REAL_TO_STRF;
		REAL_TO_STRF := CONCAT('0', st_tmp);
	END_FOR;
	IF n > 0 THEN REAL_TO_STRF := INSERT(REAL_TO_STRF, D, LEN(REAL_TO_STRF) - N); END_IF;
	IF in < 0.0 THEN st_tmp := REAL_TO_STRF; REAL_TO_STRF := CONCAT('-', st_tmp); END_IF;

END_FUNCTION_BLOCK

PROGRAM program0

	VAR
		IN :	REAL;
		N :	INT;
		D :	STRING;

        REAL_TO_STRF :	STRING;
		func_block : REAL_TO_STRF_Block;
	END_VAR
		func_block.IN := IN;
		func_block.N := N;
		func_block.D := D;
		func_block();
		REAL_TO_STRF := func_block.REAL_TO_STRF;

END_PROGRAM

CONFIGURATION Config0

	RESOURCE Res0 ON PLC
		TASK task0(INTERVAL := T#20ms,PRIORITY := 0);
		PROGRAM instance0 WITH task0 : program0;
	END_RESOURCE

END_CONFIGURATION

(* ---- 452-MESSAGE_4R.ST ---- *)
FUNCTION INC1:INT

	VAR_INPUT
		X :	INT;
		N :	INT;
	END_VAR

	IF X >= N - 1 THEN
		INC1 := 0;
	ELSE
		INC1 := X + 1;
	END_IF;
END_FUNCTION

FUNCTION_BLOCK MESSAGE_4R_Block

	VAR_INPUT
		M0 :	STRING;
		M1 :	STRING;
		M2 :	STRING;
		M3 :	STRING;
		MM :	INT := 3;
		ENQ :	BOOL := TRUE;
		CLK :	BOOL := TRUE;
		T1 :	TIME := T#3s;
	END_VAR

	VAR_OUTPUT
		MX :	STRING;
		MN :	INT;
		TR :	BOOL;
	END_VAR

	VAR
		timer :	TON;
		edge :	BOOL;
	END_VAR

	TR := FALSE;
	IF ENQ THEN
		IF (NOT edge AND clk) OR timer.q THEN
				MN := INC1(MN, MM);
				TR := TRUE;
				timer(in := FALSE);
				CASE MN OF
					0 : MX := M0;
					1 : MX := M1;
					2 : MX := M2;
					3 : MX := M3;
				END_CASE;
		END_IF;
		edge := clk;
		timer( in := CLK, pt := T1);
	ELSE
		MX := '';
		MN := 0;
	END_IF;

END_FUNCTION_BLOCK

PROGRAM program0

	VAR
		M0 :	STRING;
		M1 :	STRING;
		M2 :	STRING;
		M3 :	STRING;
		MM :	INT;
		ENQ :	BOOL;
		CLK :	BOOL;
		T1 :	TIME;

		MX :	STRING;
		MN :	INT;
		TR :	BOOL;

		func_block : MESSAGE_4R_Block;
	END_VAR

	func_block.M0 := M0;
	func_block.M1 := M1;
	func_block.M2 := M2;
	func_block.M3 := M3;
	func_block.MM := MM;
	func_block.ENQ := ENQ;
	func_block.CLK := CLK;
	func_block.T1 := T1;

	func_block();

	MX := func_block.MX;
	MN := func_block.MN;
	TR := func_block.TR;

END_PROGRAM

CONFIGURATION Config0

	RESOURCE Res0 ON PLC
		TASK task0(INTERVAL := T#20ms,PRIORITY := 0);
		PROGRAM instance0 WITH task0 : program0;
	END_RESOURCE

END_CONFIGURATION

(* ---- 453-BASE64_DECODE_STREAM.ST ---- *)
TYPE
  oscat_aB0_47	: ARRAY [0..47]	OF BYTE;
  oscat_aB0_63	: ARRAY [0..63]	OF BYTE;
END_TYPE

FUNCTION_BLOCK BASE64_DECODE_STREAM
	VAR_IN_OUT
		BUF1 :	oscat_aB0_63;
		BUF2 :	oscat_aB0_47;
	END_VAR

	VAR_INPUT
		SIZE1 :	INT;
	END_VAR

	VAR_OUTPUT
		SIZE2 :	INT;
	END_VAR

	VAR
		a :	INT;
		b :	WORD;
		o :	INT;
		off :	INT;
		i1 :	INT;
		i2 :	INT;
		c :	INT;
	END_VAR

	IF SIZE1 <= 0 THEN SIZE2 := 0; RETURN; END_IF;
	c := SIZE1 - 1;
	i2 := 0;
	a := 0;
	b := WORD#0;
	FOR i1 := 0 TO c DO
		o := BYTE_TO_INT(BUF1[i1]);
		IF o = 61  (* = *) THEN EXIT;
		ELSIF o > 96 (* a-z *) THEN off := 71;
		ELSIF o > 64 (* A-Z *) THEN off := 65;
		ELSIF o > 47 (* 0-9 *) THEN off := -4;
		ELSIF o = 43 (* + *) THEN off := -19;
		ELSIF o = 47 (* / *) THEN off := -16;
		END_IF;
		b := SHL(b,6) OR INT_TO_WORD(o - off);
		a := a + 6;
		IF a >= 8 THEN
			a := a - 8;
			BUF2[i2] := WORD_TO_BYTE(SHR(b,a));
			i2 := i2 + 1;
			b := b AND NOT SHL(WORD#16#FFFF,a);
		END_IF;
	END_FOR;
	SIZE2 := i2;
END_FUNCTION_BLOCK

PROGRAM program0
  VAR
	BUF1  :	oscat_aB0_63;
	BUF2  :	oscat_aB0_47;

	SIZE1 :	INT;

	SIZE2 :	INT;
	func_block : BASE64_DECODE_STREAM;
  END_VAR
	func_block.BUF1 :=BUF1 ;
	func_block.BUF2 :=BUF2 ;
	func_block.SIZE1:=SIZE1;
	func_block();
	BUF1 := func_block.BUF1;
	BUF2 := func_block.BUF2;
	SIZE2 := func_block.SIZE2;
END_PROGRAM

CONFIGURATION Config0
  RESOURCE Res0 ON PLC
    TASK task0(INTERVAL := T#20ms,PRIORITY := 0);
    PROGRAM instance0 WITH task0 : program0;
  END_RESOURCE
END_CONFIGURATION

(* ---- 456-SHR_8UDE.ST ---- *)
FUNCTION_BLOCK SHR_8UDE_Block

	VAR_INPUT
		SET :	BOOL;
		D0 :	BOOL;
		D7 :	BOOL;
		CLK :	BOOL;
		DN :	BOOL;
		RST :	BOOL;
	END_VAR

	VAR_OUTPUT
		Q0 :	BOOL;
		Q1 :	BOOL;
		Q2 :	BOOL;
		Q3 :	BOOL;
		Q4 :	BOOL;
		Q5 :	BOOL;
		Q6 :	BOOL;
		Q7 :	BOOL;
	END_VAR

	VAR
		trig :	R_TRIG;
	END_VAR

	trig(clk := clk);

	IF set OR rst THEN
		Q0 := NOT RST;
		Q1 := Q0;
		Q2 := Q0;
		Q3 := Q0;
		Q4 := Q0;
		Q5 := Q0;
		Q6 := Q0;
		Q7 := Q0;
	ELSIF trig.Q THEN
		IF dn THEN
			Q0 := Q1;
			Q1 := Q2;
			Q2 := Q3;
			Q3 := Q4;
			Q4 := Q5;
			Q5 := Q6;
			Q6 := Q7;
			Q7 := D7;
		ELSE
			Q7 := Q6;
			Q6 := Q5;
			Q5 := Q4;
			Q4 := Q3;
			Q3 := Q2;
			Q2 := Q1;
			Q1 := Q0;
			Q0 := D0;
		END_IF;
	END_IF;

END_FUNCTION_BLOCK

PROGRAM program0
	VAR
		SET :	BOOL;
		D0 :	BOOL;
		D7 :	BOOL;
		CLK :	BOOL;
		DN :	BOOL;
		RST :	BOOL;
		Q0 :	BOOL;
		Q1 :	BOOL;
		Q2 :	BOOL;
		Q3 :	BOOL;
		Q4 :	BOOL;
		Q5 :	BOOL;
		Q6 :	BOOL;
		Q7 :	BOOL;
		func_block : SHR_8UDE_Block;
  	END_VAR
	func_block.SET  :=SET;
	func_block.D0  :=D0;
	func_block.D7  :=D7;
	func_block.CLK  :=CLK;
	func_block.DN  :=DN;
	func_block.RST  :=RST;
	func_block();
	Q0  := func_block.Q0;
	Q1  := func_block.Q1;
	Q2  := func_block.Q2;
	Q3  := func_block.Q3;
	Q4  := func_block.Q4;
	Q5  := func_block.Q5;
	Q6  := func_block.Q6;
	Q7  := func_block.Q7;
END_PROGRAM

CONFIGURATION Config0
	RESOURCE Res0 ON PLC
		TASK task0(INTERVAL := T#20ms,PRIORITY := 0);
		PROGRAM instance0 WITH task0 : program0;
	END_RESOURCE
END_CONFIGURATION

(* ---- 457-TELNET_LOG.ST ---- *)
FUNCTION_BLOCK TELNET_LOG

	VAR_INPUT
		ENABLE :	BOOL;
		OPTION :	BYTE := BYTE#2#1000_1100;
		PORT :	WORD := WORD#23;
	END_VAR

	VAR_OUTPUT
		READY :	BOOL;
	END_VAR

	VAR_IN_OUT
		IP_C :	oscat_IP_C;
		S_BUF :	oscat_NETWORK_BUFFER;
		LOG_CL :	us_LOG_CONTROL;
	END_VAR

	VAR
		TELNET_PRINT :	TELNET_PRINT;
		done :	BOOL;
		init :	BOOL;
		watchdog :	TON;
		ci :	INT;
		pi :	INT;
		pi_last :	INT;
		send :	BOOL;
	END_VAR

	IF NOT init THEN
		init := TRUE;
		IF OPTION > BYTE#0 THEN
			TELNET_PRINT.OPTION := OPTION;
		END_IF;
		IF PORT > WORD#0 THEN
			TELNET_PRINT.PORT := PORT;
		END_IF;
		WATCHDOG.PT := T#1ms;
	END_IF;

	WATCHDOG(IN:=FALSE);

	ci := LOG_CL.IDX;

	IF IP_C.C_STATE = BYTE#1 THEN
		pi := 0;
		init := FALSE;
	END_IF;

	REPEAT
		IF pi <> ci AND IP_C.C_STATE > BYTE#127 THEN
			IF pi = 0 AND LOG_CL.RING_MODE THEN pi := ci; END_IF;
			pi_last := pi;
			pi := pi + 1;
			IF pi > LOG_CL.SIZE THEN pi := 1; END_IF;
			SEND := TRUE;
		ELSE
			SEND := FALSE;
		END_IF;

		TELNET_PRINT(	IP_C := IP_C,
						S_BUF := S_BUF,
						ENABLE := ENABLE,
						SEND := SEND,
						TEXT := LOG_CL.MSG[pi],
						BACK_COLOR := DWORD_TO_BYTE(SHL(LOG_CL.MSG_OPTION[pi],8)),
						FRONT_COLOR := DWORD_TO_BYTE(LOG_CL.MSG_OPTION[pi] ));
		READY := TELNET_PRINT.READY;
		done  := TELNET_PRINT.DONE;
		IP_C  := TELNET_PRINT.IP_C;
		S_BUF := TELNET_PRINT.S_BUF;

		IF SEND AND NOT done THEN
			pi := pi_last;
		END_IF;

		WATCHDOG(IN:=TRUE);

	UNTIL (WATCHDOG.Q OR NOT done )
	END_REPEAT;

END_FUNCTION_BLOCK

(* ---- 458-IRTRANS_RCV_4.ST ---- *)
FUNCTION_BLOCK IRTRANS_RCV_4_Block

	VAR_INPUT
		CMD :	BOOL;
	END_VAR

	VAR_IN_OUT
		DEV :	STRING;
		KEY :	STRING;
	END_VAR

	VAR_INPUT
		DEV_CODE :	STRING;
		KEY_CODE_0 :	STRING;
		KEY_CODE_1 :	STRING;
		KEY_CODE_2 :	STRING;
		KEY_CODE_3 :	STRING;
	END_VAR

	VAR_OUTPUT
		Q0 :	BOOL;
		Q1 :	BOOL;
		Q2 :	BOOL;
		Q3 :	BOOL;
	END_VAR

	VAR
		decode :	BOOL;
	END_VAR

	decode := cmd AND EQ_STRING(dev_code,dev);

	Q0 := EQ_STRING(key,key_code_0) AND decode;
	Q1 := EQ_STRING(key,key_code_1) AND decode;
	Q2 := EQ_STRING(key,key_code_2) AND decode;
	Q3 := EQ_STRING(key,key_code_3) AND decode;

END_FUNCTION_BLOCK

PROGRAM program0
	VAR
		CMD :	BOOL;
		DEV :	STRING;
		KEY :	STRING;
		DEV_CODE :	STRING;
		KEY_CODE_0 :	STRING;
		KEY_CODE_1 :	STRING;
		KEY_CODE_2 :	STRING;
		KEY_CODE_3 :	STRING;
		Q0 :	BOOL;
		Q1 :	BOOL;
		Q2 :	BOOL;
		Q3 :	BOOL;

		func_block : IRTRANS_RCV_4_Block;
	END_VAR
	func_block.CMD := CMD;
	func_block.DEV := DEV;
	func_block.KEY := KEY;
	func_block.DEV_CODE := DEV_CODE;
	func_block.KEY_CODE_0 := KEY_CODE_0;
	func_block.KEY_CODE_1 := KEY_CODE_1;
	func_block.KEY_CODE_2 := KEY_CODE_2;
	func_block.KEY_CODE_3 := KEY_CODE_3;

	func_block();
	DEV  := func_block.DEV;
	KEY  := func_block.KEY;
	Q0  := func_block.Q0;
	Q1  := func_block.Q1;
	Q2  := func_block.Q2;
	Q3  := func_block.Q3;

END_PROGRAM

CONFIGURATION Config0

  	RESOURCE Res0 ON PLC
    	TASK task0(INTERVAL := T#20ms,PRIORITY := 0);
    	PROGRAM instance0 WITH task0 : program0;
  	END_RESOURCE

END_CONFIGURATION

(* ---- 459-LENGTH.ST ---- *)
FUNCTION_BLOCK LENGTH_Block

	VAR_INPUT
		M :	REAL;
		P :	REAL;
		IN :	REAL;
		FT :	REAL;
		YD :	REAL;
		MILE :	REAL;
		SM :	REAL;
		FM :	REAL;
	END_VAR

	VAR_OUTPUT
		YM :	REAL;
		YP :	REAL;
		YIN :	REAL;
		YFT :	REAL;
		YYD :	REAL;
		YMILE :	REAL;
		YSM :	REAL;
		YFM :	REAL;
	END_VAR

	Ym :=	m
			+ p * 0.000376065
			+ in * 0.0254
			+ ft * 0.3048
			+ yd * 0.9144
			+ mile * 1609.344
			+ sm * 1852.0
			+ fm * 1.829;
	Yp := Ym * 2659.11478068951;
	Yin := Ym * 39.37007874016;
	Yft := Ym * 3.28083989501;
	Yyd := Ym * 1.09361329834;
	Ymile := Ym * 0.00062137119;
	Ysm := Ym * 0.00053995680;
	Yfm := Ym * 0.54674685621;

END_FUNCTION_BLOCK

PROGRAM program0

	VAR
		M :	REAL;
		P :	REAL;
		IN :	REAL;
		FT :	REAL;
		YD :	REAL;
		MILE :	REAL;
		SM :	REAL;
		FM :	REAL;

		YM :	REAL;
		YP :	REAL;
		YIN :	REAL;
		YFT :	REAL;
		YYD :	REAL;
		YMILE :	REAL;
		YSM :	REAL;
		YFM :	REAL;

		func_block : LENGTH_Block;
	END_VAR
	func_block.M := M;
	func_block.P := P;
	func_block.IN := IN;
	func_block.FT := FT;
	func_block.YD := YD;
	func_block.MILE := MILE;
	func_block.SM := SM;
	func_block.FM := FM;

	func_block();

	YM := func_block.YM;
	YP := func_block.YP;
	YIN := func_block.YIN;
	YFT := func_block.YFT;
	YYD := func_block.YYD;
	YMILE := func_block.YMILE;
	YSM := func_block.YSM;
	YFM := func_block.YFM;

END_PROGRAM

CONFIGURATION Config0

	RESOURCE Res0 ON PLC
		TASK task0(INTERVAL := T#20ms,PRIORITY := 0);
		PROGRAM instance0 WITH task0 : program0;
	END_RESOURCE

END_CONFIGURATION

(* ---- 460-LOG_MSG_80.ST ---- *)
FUNCTION_BLOCK LOG_MSG_80
  VAR_EXTERNAL
    LOG_CL_80 :	us_LOG_CONTROL_80;
  END_VAR

  VAR
    FB_PRINT_SF_80 :	PRINT_SF_80;
  END_VAR

  VAR
    idx :	INT;
  END_VAR

  IF DWORD_TO_BYTE(SHL(LOG_CL_80.NEW_MSG_OPTION,16)) > LOG_CL_80.LEVEL THEN RETURN; END_IF;
  LOG_CL_80.SIZE := 400;

  FB_PRINT_SF_80.PRINTF_DATA := LOG_CL_80.PRINTF;
  FB_PRINT_SF_80.STR := LOG_CL_80.NEW_MSG;
  FB_PRINT_SF_80();
  LOG_CL_80.NEW_MSG := FB_PRINT_SF_80.STR;
  LOG_CL_80.PRINTF := FB_PRINT_SF_80.PRINTF_DATA;

  IF LOG_CL_80.RESET THEN
    LOG_CL_80.RESET := FALSE;
    LOG_CL_80.RING_MODE := FALSE;
    LOG_CL_80.IDX := 0;
    LOG_CL_80.UPDATE_COUNT := LOG_CL_80.UPDATE_COUNT + UINT#1;
  END_IF;

  IF LEN(LOG_CL_80.NEW_MSG) > 0 THEN
    IF (LOG_CL_80.IDX >= LOG_CL_80.SIZE) THEN
      LOG_CL_80.RING_MODE := TRUE;
      LOG_CL_80.IDX := 0;
    END_IF;

    LOG_CL_80.UPDATE_COUNT := LOG_CL_80.UPDATE_COUNT + UINT#1;
    LOG_CL_80.IDX := LOG_CL_80.IDX + INT#1;
    idx := LOG_CL_80.IDX;
    LOG_CL_80.MSG[idx] := LOG_CL_80.NEW_MSG;
    LOG_CL_80.MSG_OPTION[idx] := LOG_CL_80.NEW_MSG_OPTION;
    LOG_CL_80.NEW_MSG := '';
  END_IF;
END_FUNCTION_BLOCK

PROGRAM program0
	VAR
		STR :	oscat_STRING80;
		LOG_MSG_80_R :	DWORD;
		func_block : LOG_MSG_80;
	END_VAR

	func_block.STR := STR;
	func_block();
	LOG_MSG_80_R  := func_block.LOG_MSG_80;
END_PROGRAM

CONFIGURATION Config0
  	RESOURCE Res0 ON PLC
    	TASK task0(INTERVAL := T#20ms,PRIORITY := 0);
    	PROGRAM instance0 WITH task0 : program0;
  	END_RESOURCE
END_CONFIGURATION

(* ---- 461-CONTROL_SET1.ST ---- *)
FUNCTION_BLOCK CONTROL_SET1_Block
	VAR_INPUT
		KT :	REAL;
		TT :	REAL;
		PI :	BOOL;
		PIDD :	BOOL;
		P_K :	REAL := 0.5;
		PI_K :	REAL := 0.45;
		PI_TN :	REAL := 0.83;
		PIDD_K :	REAL := 0.6;
		PIDD_TN :	REAL := 0.5;
		PIDD_TV :	REAL := 0.125;
	END_VAR

	VAR_OUTPUT
		KP :	REAL;
		TN :	REAL;
		TV :	REAL;
		KI :	REAL;
		KD :	REAL;
	END_VAR

	IF pi AND PIDD THEN
		KP := 0.0;
		TN := 0.0;
		TV := 0.0;
	ELSIF PIDD THEN
		KP := PIDD_K * Kt;
		TN := PIDD_TN * Tt;
		TV := PIDD_TV * Tt;
	ELSIF PI THEN
		KP := PI_K * Kt;
		TN := PI_TN * Tt;
	ELSE
		KP := P_K * Kt;
	END_IF;
	IF tn > 0.0 THEN KI := KP / TN; ELSE KI := 0.0; END_IF;
	KD := KP * TV;
END_FUNCTION_BLOCK

PROGRAM program0
  VAR
	KT :REAL;
	TT :REAL;
	PI :BOOL;
	PIDD :BOOL;
	P_K :REAL ;
	PI_K :REAL ;
	PI_TN :REAL ;
	PIDD_K :REAL ;
	PIDD_TN :REAL ;
	PIDD_TV :REAL ;
	KP :REAL;
	TN :REAL;
	TV :REAL;
	KI :REAL;
	KD :REAL;
	func_block : CONTROL_SET1_Block;
  END_VAR
	func_block.KT   :=KT  ;
	func_block.TT   :=TT  ;
	func_block.PI   :=PI  ;
	func_block.PIDD   :=PIDD  ;
	func_block.P_K   :=P_K  ;
	func_block.PI_K   :=PI_K  ;
	func_block.PI_TN   :=PI_TN  ;
	func_block.PIDD_K   :=PIDD_K  ;
	func_block.PIDD_TN   :=PIDD_TN  ;
	func_block.PIDD_TV   :=PIDD_TV  ;
	func_block();
	KP := func_block.KP ;
	TN := func_block.TN ;
	TV := func_block.TV ;
	KI := func_block.KI ;
	KD := func_block.KD ;
END_PROGRAM

CONFIGURATION Config0
  RESOURCE Res0 ON PLC
    TASK task0(INTERVAL := T#20ms,PRIORITY := 0);
    PROGRAM instance0 WITH task0 : program0;
  END_RESOURCE
END_CONFIGURATION

(* ---- 462-SDT_TO_DATE.ST ---- *)
TYPE oscat_SDT :
	STRUCT
		YEAR : INT;
		MONTH : INT;
		DAY : INT;
		WEEKDAY : INT;
		HOUR : INT;
		MINUTE : INT;
		SECOND : INT;
		MS : INT;
	END_STRUCT;
END_TYPE

FUNCTION _INT_TO_UDINT:UDINT
	VAR_INPUT
		IN :	INT;
	END_VAR

	_INT_TO_UDINT := DINT_TO_UDINT(INT_TO_DINT(IN));
END_FUNCTION

FUNCTION SET_DATE:UDINT

	VAR_INPUT
		YEAR :	INT;
		MONTH :	INT;
		DAY :	INT;
	END_VAR

	VAR
		count :	INT;
	END_VAR

	IF month > 2 THEN
		count := (month - 1) * 30;
		IF month > 7 THEN
			count := count + DWORD_TO_INT(SHR(DINT_TO_DWORD(INT_TO_DINT(month) - INT_TO_DINT(3)),1));
		ELSE
			count := count + DWORD_TO_INT(SHR(DINT_TO_DWORD(INT_TO_DINT(month) - INT_TO_DINT(4)),1));
		END_IF;
		IF SHL(INT_TO_WORD(year),14) = WORD#0 THEN
			count := count + 1;
		END_IF;
	ELSE
		count := (month - 1) * 31;
	END_IF;
	SET_DATE := (_INT_TO_UDINT(count + day - 1) + DWORD_TO_UDINT(SHR(UDINT_TO_DWORD(_INT_TO_UDINT(year) * UDINT#1461 - UDINT#2878169), 2))) * UDINT#86400;

END_FUNCTION

FUNCTION_BLOCK SDT_TO_DATE_Block

	VAR_INPUT
		DTI :	oscat_SDT;
	END_VAR

	VAR_OUTPUT
		SDT_TO_DATE :	UDINT;
	END_VAR

	SDT_TO_DATE := SET_DATE(DTI.YEAR, DTI.MONTH, DTI.DAY);

END_FUNCTION_BLOCK

PROGRAM program0

	VAR
		DTI :	oscat_SDT;
		SDT_TO_DATE :	UDINT;
		func_block : SDT_TO_DATE_Block;
  	END_VAR
	func_block.DTI  :=	DTI;
	func_block();
	SDT_TO_DATE := func_block.SDT_TO_DATE;

END_PROGRAM

CONFIGURATION Config0

	RESOURCE Res0 ON PLC
		TASK task0(INTERVAL := T#20ms,PRIORITY := 0);
		PROGRAM instance0 WITH task0 : program0;
	END_RESOURCE

END_CONFIGURATION

(* ---- 463-BUFFER_COMP_NW.ST ---- *)
TYPE
  oscat_NW_BUF_LONG  : ARRAY [0..4095] OF BYTE;
END_TYPE

FUNCTION_BLOCK BUFFER_COMP_NW
	VAR_IN_OUT
		PT1 :	oscat_NW_BUF_LONG;
	END_VAR

	VAR_INPUT
		SIZE1 :	INT;
	END_VAR

	VAR_IN_OUT
		PT2 :	oscat_NW_BUF_LONG;
	END_VAR

	VAR_INPUT
		SIZE2 :	INT;
		START :	INT;
	END_VAR

	VAR_OUTPUT
		BUFFER_COMP :	INT;
	END_VAR

	VAR
		i :	INT;
		j :	INT;
		end :	INT;
		j2 :	INT;
	END_VAR

	IF SIZE2 <= SIZE1 AND SIZE1 > 0 AND SIZE2 > 0 AND START >= 0 THEN
		end := SIZE1 - SIZE2;
		FOR i := START TO end DO
			IF PT1[i] = PT2[0] THEN
				(* first character matches, now compare rest of array *)
				j := 1;
				j2 := j + i;
				WHILE j < SIZE2 DO
					IF PT2[j] <> PT1[j2] THEN EXIT; END_IF;
					j := j + 1;
					j2 := j2 + 1;
				END_WHILE;
				(* when J > size2 a match was found return the position i in buffer1 *)
				IF j = SIZE2 THEN
					BUFFER_COMP := i;
					RETURN;
				END_IF;
			END_IF;
		END_FOR;
	END_IF;
	BUFFER_COMP := -1;

END_FUNCTION_BLOCK

PROGRAM program0
  VAR
	PT1   :	oscat_NW_BUF_LONG;

	SIZE1 :	INT;

	PT2   : 	oscat_NW_BUF_LONG;

	SIZE2 :	INT;
	START :	INT;

	BUFFER_COMP :	INT;

	func_block : BUFFER_COMP_NW;
  END_VAR
	func_block.PT1  :=PT1  ;
	func_block.SIZE1:=SIZE1;
	func_block.PT2  :=PT2  ;
	func_block.SIZE2:=SIZE2;
	func_block.START:=START;
	func_block();
	BUFFER_COMP := func_block.BUFFER_COMP;
	PT1 := func_block.PT1;
	PT2 := func_block.PT2;

END_PROGRAM

CONFIGURATION Config0
  RESOURCE Res0 ON PLC
    TASK task0(INTERVAL := T#20ms,PRIORITY := 0);
    PROGRAM instance0 WITH task0 : program0;
  END_RESOURCE
END_CONFIGURATION

(* ---- 464-LAMBERT_W.ST ---- *)
FUNCTION _REAL_TO_DWORD: DWORD

  VAR_INPUT
    X :	REAL;
  END_VAR

  IF REAL_TO_DWORD(0.5) = DWORD#1 THEN
    _REAL_TO_DWORD := REAL_TO_DWORD(x);
  ELSIF X > 0.0 THEN
    _REAL_TO_DWORD := REAL_TO_DWORD(x+0.5);
  ELSIF X < 0.0 THEN
    _REAL_TO_DWORD := REAL_TO_DWORD(x-0.5);
  ELSE
    _REAL_TO_DWORD := DWORD#0;
  END_IF;
END_FUNCTION

FUNCTION_BLOCK LAMBERT_W_Block

	VAR_INPUT
		X :	REAL;
	END_VAR

	VAR_OUTPUT
		LAMBERT_W :	REAL;
	END_VAR

	VAR
		w :	REAL;
		i :	INT;
		we :	REAL;
		w1e :	REAL;
		last :	DWORD;
		ewx :	REAL;
	END_VAR

	IF x < -0.367879441171442 THEN
		LAMBERT_W := -1000.0;
		RETURN;
	(* return 0 if x = 0 *)
	ELSIF x = 0.0 THEN
		RETURN;
	(* first an estimate is calculated *)
	ELSIF x <= 500.0 THEN
		w := LN(x + 1.0);
		w := 0.665 * (1.0 + 0.0195 * w) * w + 0.04;
	ELSE
		w := LN(x - 4.0) - (1.0 - 1.0/LN(x)) * LN(LN(x));
	END_IF;
	(* use estimate to calculate exact result *)
	FOR i := 0 TO 5 DO
		ewx := EXP(w);
		we := w * ewx - x;
		w1e := (w+1.0) * ewx;
		last := _REAL_TO_DWORD(w) AND DWORD#16#FFFF_FFFC;
		w := w - (we / (w1e - (w+2.0) * we / (2.0 * w + 2.0)));
		IF (_REAL_TO_DWORD(w) AND DWORD#16#FFFF_FFFC) = last THEN EXIT; END_IF;
	END_FOR;
	LAMBERT_W := w;

END_FUNCTION_BLOCK

PROGRAM program0

	VAR
		X :	REAL;
		LAMBERT_W :	REAL;
		func_block : LAMBERT_W_Block;
	END_VAR
	func_block.X := X;
	func_block();
	LAMBERT_W := func_block.LAMBERT_W;

END_PROGRAM

CONFIGURATION Config0

	RESOURCE Res0 ON PLC
		TASK task0(INTERVAL := T#20ms,PRIORITY := 0);
		PROGRAM instance0 WITH task0 : program0;
	END_RESOURCE

END_CONFIGURATION

(* ---- 465-BUFFER_TO_STRING.ST ---- *)
TYPE
	oscat_arb_0_249 			  : ARRAY [0..249] 	OF BYTE;
END_TYPE

FUNCTION_BLOCK BUFFER_TO_STRING_Block
	VAR_IN_OUT
		PT  :	oscat_arb_0_249;
	END_VAR

	VAR_INPUT
		SIZE :	UINT;
		START :	UINT;
		STOP :	UINT;
	END_VAR

	VAR_OUTPUT
		BUFFER_TO_STRING :	STRING;
	END_VAR

	VAR
		sta :	UINT;
		stp :	UINT;
		size2 :	UINT;
		i :	INT;
		BUF_TO_STRING :	BUF_TO_STRING;
	END_VAR

	sta := MIN(START, SIZE - UINT#1);
	stp := STOP;
	IF stp - sta + UINT#1 > UINT#250 THEN
		stp := sta + UINT#250 - UINT#1;
	END_IF;
	stp := MIN(stp, SIZE - UINT#1);
	size2 := stp - sta + UINT#1;
	IF size2 > UINT#0 THEN
		FOR i := 0 TO 1 DO
			BUF_TO_STRING.REQ := i > 0;
			BUF_TO_STRING.BUF_FORMAT := TRUE;
			BUF_TO_STRING.BUF_OFFS := UINT_TO_DINT(START);
			BUF_TO_STRING.BUF_CNT := UINT_TO_DINT(size2);
			BUF_TO_STRING.BUFFER := pt;
			BUF_TO_STRING.DST := BUFFER_TO_STRING;
			BUF_TO_STRING();
			pt := BUF_TO_STRING.BUFFER;
			BUFFER_TO_STRING := BUF_TO_STRING.DST;
		END_FOR;
	ELSE
		BUFFER_TO_STRING :='';
	END_IF;
END_FUNCTION_BLOCK

PROGRAM program0
  VAR
    LocalVar0 : oscat_arb_0_249;
    LocalVar1 : UINT;
	LocalVar2 : UINT;
	LocalVar3 : UINT;
	LocalOUT  : INT;
	func_block : BUFFER_TO_STRING_Block;
  END_VAR
	func_block.PT  := LocalVar0;
	func_block.SIZE := LocalVar1;
	func_block.START := LocalVar2;
	func_block.STOP := LocalVar3;
	func_block();
	LocalOUT := func_block.BUFFER_TO_STRING;
	LocalVar0 := func_block.PT;

END_PROGRAM

CONFIGURATION Config0
  RESOURCE Res0 ON PLC
    TASK task0(INTERVAL := T#20ms,PRIORITY := 0);
    PROGRAM instance0 WITH task0 : program0;
  END_RESOURCE
END_CONFIGURATION

(* ---- 466-MESSAGE_8.ST ---- *)
FUNCTION_BLOCK MESSAGE_8_Block

	VAR_INPUT
		IN1 :	BOOL;
		IN2 :	BOOL;
		IN3 :	BOOL;
		IN4 :	BOOL;
		IN5 :	BOOL;
		IN6 :	BOOL;
		IN7 :	BOOL;
		IN8 :	BOOL;
		S1 :	STRING;
		S2 :	STRING;
		S3 :	STRING;
		S4 :	STRING;
		S5 :	STRING;
		S6 :	STRING;
		S7 :	STRING;
		S8 :	STRING;
	END_VAR

	VAR_OUTPUT
		M :	STRING;
	END_VAR

	IF in1 THEN
		M := S1;
	ELSIF in2 THEN
		M := S2;
	ELSIF in3 THEN
		M := S3;
	ELSIF in4 THEN
		M := S4;
	ELSIF in5 THEN
		M := S5;
	ELSIF in6 THEN
		M := S6;
	ELSIF in7 THEN
		M := S7;
	ELSIF in8 THEN
		M := S8;
	ELSE
		M := '';
	END_IF;

END_FUNCTION_BLOCK

PROGRAM program0

	VAR
		IN1 :	BOOL;
		IN2 :	BOOL;
		IN3 :	BOOL;
		IN4 :	BOOL;
		IN5 :	BOOL;
		IN6 :	BOOL;
		IN7 :	BOOL;
		IN8 :	BOOL;
		S1 :	STRING;
		S2 :	STRING;
		S3 :	STRING;
		S4 :	STRING;
		S5 :	STRING;
		S6 :	STRING;
		S7 :	STRING;
		S8 :	STRING;

		M :	STRING;

		func_block : MESSAGE_8_Block;
	END_VAR

	func_block.IN1 := IN1;
	func_block.IN2 := IN2;
	func_block.IN3 := IN3;
	func_block.IN4 := IN4;
	func_block.IN5 := IN5;
	func_block.IN6 := IN6;
	func_block.IN7 := IN7;
	func_block.IN8 := IN8;
	func_block.S1 := S1;
	func_block.S2 := S2;
	func_block.S3 := S3;
	func_block.S4 := S4;
	func_block.S5 := S5;
	func_block.S6 := S6;
	func_block.S7 := S7;
	func_block.S8 := S8;

	func_block();

	M  := func_block.M;

END_PROGRAM

CONFIGURATION Config0

	VAR_GLOBAL
		PLC_TICKS_PER_SEC :	INT;
		PLC_SYS_TICK_CNT :	DINT;
	END_VAR

	RESOURCE Res0 ON PLC
		TASK task0(INTERVAL := T#20ms,PRIORITY := 0);
		PROGRAM instance0 WITH task0 : program0;
	END_RESOURCE

END_CONFIGURATION

(* ---- 467-T_PLC_MS.ST ---- *)
FUNCTION_BLOCK T_PLC_MS_block

	VAR_OUTPUT
		T_PLC_MS :	UDINT;
	END_VAR

	VAR_EXTERNAL
		PLC_TICKS_PER_SEC :	INT;
		PLC_SYS_TICK_CNT :	DINT;
	END_VAR

	VAR
		debug :	BOOL;(*Debug-Mode ON / OFF*)
		N :	INT;(*Debug-Faktor*)
		Offset :	UDINT;(*Debug-Offset*)
		temp :	DWORD := DWORD#1;(*Debug-Offset*)
		mode :	BOOL;(*modus*)
		faktor :	UDINT;(*Systemtakt-Faktor*)
		init :	BOOL;
		v_plc_ticks_per_sec :	UDINT;
		base :	UDINT := UDINT#1000;
	END_VAR

	IF init = FALSE THEN
		v_plc_ticks_per_sec := INT_TO_UDINT(PLC_TICKS_PER_SEC);
		IF v_plc_ticks_per_sec = UDINT#1024 THEN
			faktor := UDINT#1;
			mode := FALSE;
		ELSIF v_plc_ticks_per_sec > UDINT#0 THEN
			IF v_plc_ticks_per_sec <= base THEN
				faktor := base / v_plc_ticks_per_sec;
				mode := FALSE;
			ELSE
				faktor := v_plc_ticks_per_sec / base;
				mode := TRUE;
			END_IF;
		ELSE
			faktor := UDINT#1;
		END_IF;
		init := TRUE;
	END_IF;

	IF mode THEN
		T_PLC_MS := DINT_TO_UDINT(PLC_SYS_TICK_CNT) / faktor;
	ELSE
		T_PLC_MS := DINT_TO_UDINT(PLC_SYS_TICK_CNT) * faktor;
	END_IF;

	IF debug THEN
		T_PLC_MS := (DWORD_TO_UDINT(SHL(UDINT_TO_DWORD(T_PLC_MS),N) OR SHL(temp,N)) - UDINT#1) + Offset;
	END_IF;

END_FUNCTION_BLOCK

PROGRAM program0

	VAR
		LocalOUT  : UDINT;
		func_block : T_PLC_MS_block;
  	END_VAR

	func_block();
	LocalOUT := func_block.T_PLC_MS;

END_PROGRAM

CONFIGURATION Config0

	VAR_GLOBAL
		PLC_TICKS_PER_SEC :	INT;
		PLC_SYS_TICK_CNT :	DINT;
	END_VAR

  	RESOURCE Res0 ON PLC
    	TASK task0(INTERVAL := T#20ms,PRIORITY := 0);
    	PROGRAM instance0 WITH task0 : program0;
  	END_RESOURCE

END_CONFIGURATION

(* ---- 469-FT_AVG.ST ---- *)
TYPE
	oscat_delay_buf             : ARRAY [0..31]   OF REAL;
END_TYPE

FUNCTION INC1:INT

	VAR_INPUT
		X :	INT;
		N :	INT;
	END_VAR

	IF X >= N - 1 THEN
		INC1 := 0;
	ELSE
		INC1 := X + 1;
	END_IF;
END_FUNCTION

FUNCTION_BLOCK DELAY

	VAR_INPUT
		IN :	REAL;
		N :	INT;
		RST :	BOOL;
	END_VAR

	VAR_OUTPUT
		OUT :	REAL;
	END_VAR

	VAR
		buf :	oscat_delay_buf;
		i :	INT;
		init :	BOOL;
		stop :	INT;
	END_VAR

	stop := LIMIT(0,N,32) - 1;
	IF rst OR NOT init THEN
		init := TRUE;
		FOR i := 0 TO stop DO buf[i] := in; END_FOR;
		out := in;
		i := 0;
	ELSIF stop < 0 THEN
		out := in;
	ELSE
		out := buf[i];
		buf[i] := in;
		i := INC1(i, N);
	END_IF;

END_FUNCTION_BLOCK

FUNCTION_BLOCK FT_AVG

	VAR_INPUT
		IN :	REAL;
		E :	BOOL := TRUE;
		N :	INT := INT#32;
		RST :	BOOL;
	END_VAR

	VAR_OUTPUT
		AVG :	REAL;
	END_VAR

	VAR
		buff :	delay;
		i :	INT;
		init :	BOOL;
	END_VAR

	buff.N := LIMIT(0, N, 32);

	IF NOT init OR rst THEN
		FOR i := 1 TO N DO
			buff(in := in);
		END_FOR;
		avg := in;
		init := TRUE;
	ELSIF E THEN
		buff(in := in);
		avg := avg + (in - buff.out ) / INT_TO_REAL(N);
	END_IF;

END_FUNCTION_BLOCK

PROGRAM program0
  VAR
		IN  :	REAL;
		E   :	BOOL;
		N   :	INT;
		RST :	BOOL;

		AVG :	REAL;

	func_block : FT_AVG;
  END_VAR
	func_block.IN :=IN ;
	func_block.E  :=E  ;
	func_block.N  :=N  ;
	func_block.RST:=RST;
	func_block();
	AVG := func_block.AVG;
END_PROGRAM

CONFIGURATION Config0
  RESOURCE Res0 ON PLC
    TASK task0(INTERVAL := T#20ms,PRIORITY := 0);
    PROGRAM instance0 WITH task0 : program0;
  END_RESOURCE
END_CONFIGURATION

(* ---- 471-REPLACE_ALL.ST ---- *)
FUNCTION_BLOCK FINDP_Block

	VAR_INPUT
		STR :	STRING;
		SRC :	STRING;
		POS :	INT;
	END_VAR

	VAR_OUTPUT
		FINDP :	INT;
	END_VAR

	VAR
		i :	INT;
		ls :	INT;
		lx :	INT;
		stp :	INT;
		st_tmp :	STRING;
	END_VAR

	ls := LEN(str);
	lx := LEN(src);
	IF ls < lx OR lx = 0 THEN RETURN; END_IF;
	stp := ls - lx + 1;
	FOR i := MAX(pos,1) TO stp DO
		st_tmp := MID(str,lx,i);
		IF EQ_STRING(st_tmp,src) THEN
			FINDP := i;
			RETURN;
		END_IF;
	END_FOR;
	FINDP := 0;

END_FUNCTION_BLOCK

FUNCTION_BLOCK REPLACE_ALL_Block

	VAR_INPUT
		STR :	STRING;
		SRC :	STRING;
		REP :	STRING;
	END_VAR

	VAR_OUTPUT
		REPLACE_ALL :	STRING;
	END_VAR

	VAR
		pos :	INT;
		lp :	INT;
		lx :	INT;
		FINDP :	FINDP_Block;
		st_tmp :	STRING;
	END_VAR

	REPLACE_ALL := str;
	lx := LEN(src);
	lp := LEN(rep);

	FINDP.str := REPLACE_ALL;
	FINDP.src := src;
	FINDP.pos := 1;
	FINDP();
	pos := FINDP.FINDP;

	WHILE pos > 0 DO
		st_tmp := REPLACE_ALL;
		REPLACE_ALL := REPLACE(st_tmp,rep,lx,pos);

		FINDP.str := REPLACE_ALL;
		FINDP.src := src;
		FINDP.pos := pos + lp;
		FINDP();
		pos := FINDP.FINDP;

	END_WHILE;

END_FUNCTION_BLOCK

PROGRAM program0

	VAR
		STR :	STRING;
		SRC :	STRING;
		REP :	STRING;

        REPLACE_ALL :	STRING;
		func_block : REPLACE_ALL_Block;
	END_VAR
		func_block.STR := STR;
		func_block.SRC := SRC;
		func_block.REP := REP;
		func_block();
		REPLACE_ALL := func_block.REPLACE_ALL;

END_PROGRAM

CONFIGURATION Config0

	RESOURCE Res0 ON PLC
		TASK task0(INTERVAL := T#20ms,PRIORITY := 0);
		PROGRAM instance0 WITH task0 : program0;
	END_RESOURCE

END_CONFIGURATION

(* ---- 472-BASE64_ENCODE_STREAM.ST ---- *)
TYPE
  oscat_aB0_47	: ARRAY [0..47]	OF BYTE;
  oscat_aB0_63	: ARRAY [0..63]	OF BYTE;
END_TYPE

FUNCTION_BLOCK BASE64_ENCODE_STREAM

	VAR_IN_OUT
		BUF1 :	oscat_aB0_47;
		BUF2 :	oscat_aB0_63;
	END_VAR

	VAR_INPUT
		SIZE1 :	INT;
	END_VAR

	VAR_OUTPUT
		SIZE2 :	INT;
	END_VAR

	VAR
		a :	INT;
		b :	WORD;
		i :	INT;
		i2 :	INT;
		i3 :	INT;
		c :	INT;
		BASE64 :	STRING := 'ABCDEFGHIJKLMNOPQRSTUVWXYZabcdefghijklmnopqrstuvwxyz0123456789+/';
	END_VAR

	IF SIZE1 <= 0 THEN
		SIZE2 := 0;
		RETURN;
	END_IF;
	c := SIZE1 - 1;
	i2 := 0;
	a := 0;
	b := WORD#0;
	FOR i := 0 TO c DO
		b := SHL(b,8) OR BYTE_TO_WORD(BUF1[i]);
		a := a + 8;
		WHILE a >= 6 DO
			a := a - 6;
			buf2[i2] := INT_TO_BYTE(GET_CHAR(BASE64,WORD_TO_INT(SHR(b,a)) + 1));
			i2 := i2 + 1;
			b := b AND NOT SHL(WORD#16#FFFF,a);
		END_WHILE;
	END_FOR;
	IF a > 0 THEN
		buf2[i2] := INT_TO_BYTE(GET_CHAR(BASE64,WORD_TO_INT(SHL(b,6 - a)) + 1));
		i2 := i2 + 1;
		i3 := i2 + WORD_TO_INT(NOT INT_TO_WORD(i2) AND WORD#2#11);
		FOR i := i2 TO i3 DO
			buf2[i] := BYTE#61;
		END_FOR;
		SIZE2 := i3 + 1;
	ELSE
		SIZE2 := i2;
	END_IF;

END_FUNCTION_BLOCK

PROGRAM program0
  VAR
	BUF1  :	oscat_aB0_63;
	BUF2  :	oscat_aB0_47;

	SIZE1 :	INT;

	SIZE2 :	INT;
	func_block : BASE64_ENCODE_STREAM;
  END_VAR
	func_block.BUF1 :=BUF1 ;
	func_block.BUF2 :=BUF2 ;
	func_block.SIZE1:=SIZE1;
	func_block();
	BUF1 := func_block.BUF1;
	BUF2 := func_block.BUF2;
	SIZE2 := func_block.SIZE2;
END_PROGRAM

CONFIGURATION Config0
  RESOURCE Res0 ON PLC
    TASK task0(INTERVAL := T#20ms,PRIORITY := 0);
    PROGRAM instance0 WITH task0 : program0;
  END_RESOURCE
END_CONFIGURATION

(* ---- 473-URL_DECODE.ST ---- *)
TYPE
  oscat_STRING250               : STRING;
  oscat_STRING20               : STRING;
END_TYPE

FUNCTION_BLOCK HEX_TO_DWORD_Block

	VAR_INPUT
		HEX :	oscat_STRING20;
	END_VAR

	VAR_OUTPUT
		HEX_TO_DWORD :	DWORD;
	END_VAR

	VAR
		i :	INT;
		stop :	INT;
		X :	INT;
	END_VAR

	HEX_TO_DWORD := DWORD#0;
	stop := LEN(Hex);
	FOR I := 1 TO stop DO
		x := GET_CHAR(Hex,I);
		IF X > 47 AND x < 58 THEN
			HEX_TO_DWORD := SHL_DWORD(HEX_TO_DWORD,4) OR INT_TO_DWORD (X - 48);
		ELSIF X > 64 AND X < 71 THEN
			HEX_TO_DWORD := SHL_DWORD(HEX_TO_DWORD,4) OR INT_TO_DWORD (X - 55);
		ELSIF X > 96 AND X < 103 THEN
			HEX_TO_DWORD := SHL_DWORD(HEX_TO_DWORD,4) OR INT_TO_DWORD (X - 87);
		END_IF;
	END_FOR;

END_FUNCTION_BLOCK

FUNCTION_BLOCK URL_DECODE_Block

	VAR_INPUT
		IN :	oscat_STRING250;
	END_VAR

	VAR_OUTPUT
		URL_DECODE :	oscat_STRING250;
	END_VAR

	VAR
		pos :	INT;
		new :	STRING;
		HEX_TO_DWORD :	HEX_TO_DWORD_Block;
	END_VAR

	URL_DECODE := IN;
	pos := FIND(URL_DECODE,'%');
	WHILE pos > 0 DO
		HEX_TO_DWORD(Hex:=MID(URL_DECODE,2,pos + 1));
		new := BYTE_TO_STRING(DWORD_TO_BYTE(HEX_TO_DWORD.HEX_TO_DWORD),'%c');
		URL_DECODE := REPLACE(URL_DECODE, new, 3, pos);
		pos := FIND(URL_DECODE,'%');
	END_WHILE;

END_FUNCTION_BLOCK

PROGRAM program0
	VAR
		IN :	oscat_STRING250;
		URL_DECODE :	oscat_STRING250;

		func_block : URL_DECODE_Block;
	END_VAR
	func_block.IN := IN;

	func_block();
	URL_DECODE  := func_block.URL_DECODE;
END_PROGRAM

CONFIGURATION Config0
	RESOURCE Res0 ON PLC
		TASK task0(INTERVAL := T#20ms,PRIORITY := 0);
		PROGRAM instance0 WITH task0 : program0;
	END_RESOURCE
END_CONFIGURATION

(* ---- 474-BUFFER_COMP.ST ---- *)
TYPE
	oscat_arb_0_249 			  : ARRAY [0..249] 	OF BYTE;
END_TYPE

FUNCTION_BLOCK BUFFER_COMP_Block
	VAR_IN_OUT
		PT1 :	oscat_arb_0_249;
	END_VAR

	VAR_INPUT
		SIZE1 :	INT;
	END_VAR

	VAR_IN_OUT
		PT2 :	oscat_arb_0_249;
	END_VAR

	VAR_INPUT
		SIZE2 :	INT;
		START :	INT;
	END_VAR

	VAR_OUTPUT
		BUFFER_COMP :	INT;
	END_VAR

	VAR
		i :	INT;
		j :	INT;
		end :	INT;
		j2 :	INT;
	END_VAR

	IF SIZE2 <= SIZE1 AND SIZE1 > 0 AND SIZE2 > 0 AND START >= 0 THEN
		end := SIZE1 - SIZE2;
		FOR i := START TO end DO
			IF PT1[i] = PT2[0] THEN
				(* first character matches, now compare rest of array *)
				j := 1;
				j2 := j + i;
				WHILE j < SIZE2 DO
					IF PT2[j] <> PT1[j2] THEN EXIT; END_IF;
					j := j + 1;
					j2 := j2 + 1;
				END_WHILE;
				(* when J > size2 a match was found return the position i in buffer1 *)
				IF j = SIZE2 THEN
					BUFFER_COMP := i;
					RETURN;
				END_IF;
			END_IF;
		END_FOR;
	END_IF;
	BUFFER_COMP := -1;

END_FUNCTION_BLOCK

PROGRAM program0
  VAR
    LocalVar0 : oscat_arb_0_249;
    LocalVar1 : INT;
	LocalVar2 : oscat_arb_0_249;
	LocalVar3 : INT;
	LocalVar4 : INT;
	LocalOUT  : INT;
	func_block : BUFFER_COMP_Block;
  END_VAR
	func_block.PT1  := LocalVar0;
	func_block.SIZE1 := LocalVar1;
	func_block.PT2  := LocalVar2;
	func_block.SIZE2 := LocalVar3;
	func_block.START := LocalVar4;
	func_block();
	LocalOUT := func_block.BUFFER_COMP;
	LocalVar0 := func_block.PT1;
	LocalVar2 := func_block.PT1;

END_PROGRAM

CONFIGURATION Config0
  RESOURCE Res0 ON PLC
    TASK task0(INTERVAL := T#20ms,PRIORITY := 0);
    PROGRAM instance0 WITH task0 : program0;
  END_RESOURCE
END_CONFIGURATION

(* ---- 475-CHARCODE.ST ---- *)
TYPE
  oscat_CHARNAMES	: ARRAY [1..11] OF STRING;
END_TYPE

FUNCTION_BLOCK SETUP_CHARNAMES_Block

	VAR_IN_OUT
		CHARNAMES :	oscat_CHARNAMES;
	END_VAR

	VAR
		init :	BOOL;
	END_VAR

	IF init THEN RETURN; END_IF;

	init := TRUE;

	CHARNAMES[01] := '123';
	CHARNAMES[02] := '456';
	CHARNAMES[03] := 'zgsdafasf';
	CHARNAMES[04] := 'sadfsdfa';
	CHARNAMES[05] := 'asdfdsafdfds';
	CHARNAMES[06] := 'sadfsdfsdf';
	CHARNAMES[07] := 'sfsfdfdddd';
	CHARNAMES[08] := 'dddddted';
	CHARNAMES[10] := 'wer';
	CHARNAMES[11] := 'werwer';

END_FUNCTION_BLOCK

FUNCTION_BLOCK CHARCODE_Block
	VAR_INPUT
		STR :	STRING;
	END_VAR

	VAR_OUTPUT
		CHARCODE :	BYTE;
	END_VAR

	VAR
		found :	STRING;
		search :	STRING;
		pos :	INT;
		CODE :	CODE;
		i :	INT;
		SETUP_CHARNAMES :	SETUP_CHARNAMES_Block;
		CHARNAMES :	oscat_CHARNAMES;
	END_VAR

	SETUP_CHARNAMES(CHARNAMES:=CHARNAMES);
	CHARNAMES:=SETUP_CHARNAMES.CHARNAMES;

	IF LEN(str) = 1 THEN
		CODE(STR:=STR,POS:=1);
		CHARCODE:=CODE.CODE;
	ELSIF LEN(str) > 0 THEN
		search := CONCAT('&', str);
		search := CONCAT(search, ';');
		WHILE pos = 0 AND (i < 11) DO
			i := i + 1;
			pos := FIND(CHARNAMES[i], search);
		END_WHILE;
		found := MID(CHARNAMES[i], 1, pos - 1);
		CODE(STR:=found,POS:=1);
		CHARCODE:=CODE.CODE;
	END_IF;
END_FUNCTION_BLOCK

PROGRAM program0
  VAR
	STR :	STRING;
	CHARCODE :	BYTE;
	func_block : CHARCODE_Block;
  END_VAR
	func_block.STR  :=STR ;
	func_block();
	CHARCODE := func_block.CHARCODE;
END_PROGRAM

CONFIGURATION Config0
	RESOURCE Res0 ON PLC
		TASK task0(INTERVAL := T#20ms,PRIORITY := 0);
		PROGRAM instance0 WITH task0 : program0;
	END_RESOURCE
END_CONFIGURATION

(* ---- 476-CONTROL_SET2.ST ---- *)
FUNCTION_BLOCK CONTROL_SET2
	VAR_INPUT
		KS :	REAL;
		TU :	REAL;
		TG :	REAL;
		PI :	BOOL;
		PIDD :	BOOL;
		P_K :	REAL := 1.0;
		PI_K :	REAL := 0.9;
		PI_TN :	REAL := 3.33;
		PIDD_K :	REAL := 1.2;
		PIDD_TN :	REAL := 2.0;
		PIDD_TV :	REAL := 0.5;
	END_VAR

	VAR_OUTPUT
		KP :	REAL;
		TN :	REAL;
		TV :	REAL;
		KI :	REAL;
		KD :	REAL;
	END_VAR

	VAR
		TX :	REAL;
	END_VAR

	IF TU > 0.0 AND KS > 0.0 THEN TX := TG / TU / KS; END_IF;
	IF pi AND PIDD THEN
		KP := 0.0;
		TN := 0.0;
		TV := 0.0;
	ELSIF PIDD THEN
		KP := PIDD_K * TX;
		TN := PIDD_TN * TU;
		TV := PIDD_TV * TU;
	ELSIF PI THEN
		KP := PI_K * TX;
		TN := PI_TN * TU;
	ELSE
		KP := P_K * TX;
	END_IF;

	IF TN > 0.0 THEN KI := KP / TN; ELSE KI := 0.0; END_IF;
	KD := KP * TV;

END_FUNCTION_BLOCK

PROGRAM program0
  VAR
	KS :REAL;
	TG :REAL;
	PI :BOOL;
	PIDD :BOOL;
	P_K :REAL ;
	PI_K :REAL ;
	PI_TN :REAL ;
	PIDD_K :REAL ;
	PIDD_TN :REAL ;
	PIDD_TV :REAL ;
	KP :REAL;
	TN :REAL;
	TV :REAL;
	KI :REAL;
	KD :REAL;
	func_block : CONTROL_SET2;
  END_VAR
	func_block.KS   := KS  ;
	func_block.TG   :=TG  ;
	func_block.PI   :=PI  ;
	func_block.PIDD   :=PIDD  ;
	func_block.P_K   :=P_K  ;
	func_block.PI_K   :=PI_K  ;
	func_block.PI_TN   :=PI_TN  ;
	func_block.PIDD_K   :=PIDD_K  ;
	func_block.PIDD_TN   :=PIDD_TN  ;
	func_block.PIDD_TV   :=PIDD_TV  ;
	func_block();
	KP := func_block.KP ;
	TN := func_block.TN ;
	TV := func_block.TV ;
	KI := func_block.KI ;
	KD := func_block.KD ;
END_PROGRAM

CONFIGURATION Config0
  RESOURCE Res0 ON PLC
    TASK task0(INTERVAL := T#20ms,PRIORITY := 0);
    PROGRAM instance0 WITH task0 : program0;
  END_RESOURCE
END_CONFIGURATION

(* ---- 477-DEC_8.ST ---- *)
FUNCTION BIT_LOAD_B:BYTE
	VAR_INPUT
		IN :	BYTE;
		VAL :	BOOL;
		POS :	INT;
	END_VAR

	IF VAL THEN
		BIT_LOAD_B := in OR SHL(BYTE#1,pos);
	ELSE
		BIT_LOAD_B := in AND (NOT SHL(BYTE#1,pos));
	END_IF;
END_FUNCTION

FUNCTION _BYTE_TO_INT:INT
	VAR_INPUT
		IN :	BYTE;
	END_VAR

	_BYTE_TO_INT := USINT_TO_INT(BYTE_TO_USINT(IN));
END_FUNCTION

FUNCTION_BLOCK DEC_8

	VAR_INPUT
		D :	BOOL;
		A0 :	BOOL;
		A1 :	BOOL;
		A2 :	BOOL;
	END_VAR

	VAR_OUTPUT
		Q0 :	BOOL;
		Q1 :	BOOL;
		Q2 :	BOOL;
		Q3 :	BOOL;
		Q4 :	BOOL;
		Q5 :	BOOL;
		Q6 :	BOOL;
		Q7 :	BOOL;
	END_VAR

	VAR
		X :	BYTE;
	END_VAR

	X:=BIT_LOAD_B(X,A0,0); (* X.0 := A0; *)
	X:=BIT_LOAD_B(X,A1,1); (* X.1 := A1; *)
	X:=BIT_LOAD_B(X,A2,2); (* X.2 := A2; *)

	Q0 := FALSE;
	Q1 := FALSE;
	Q2 := FALSE;
	Q3 := FALSE;
	Q4 := FALSE;
	Q5 := FALSE;
	Q6 := FALSE;
	Q7 := FALSE;

	CASE _BYTE_TO_INT(X) OF
		0 : Q0 := D;
		1 : Q1 := D;
		2 : Q2 := D;
		3 : Q3 := D;
		4 : Q4 := D;
		5 : Q5 := D;
		6 : Q6 := D;
		7 : Q7 := D;
	END_CASE;

	END_FUNCTION_BLOCK

PROGRAM program0
  VAR
	D :	BOOL;
	A0 :	BOOL;
	A1 :	BOOL;
	A2 :	BOOL;

	Q0 :	BOOL;
	Q1 :	BOOL;
	Q2 :	BOOL;
	Q3 :	BOOL;
	Q4 :	BOOL;
	Q5 :	BOOL;
	Q6 :	BOOL;
	Q7 :	BOOL;

	func_block : DEC_8;
  END_VAR
	func_block.D   := D  ;
	func_block.A0  := A0  ;
	func_block.A1  := A1  ;
	func_block.A2  := A2  ;
	func_block();
	Q0:= func_block.Q0;
	Q1:= func_block.Q1;
	Q2:= func_block.Q2;
	Q3:= func_block.Q3;
	Q4:= func_block.Q4;
	Q5:= func_block.Q5;
	Q6:= func_block.Q6;
	Q7:= func_block.Q7;
END_PROGRAM

CONFIGURATION Config0
  RESOURCE Res0 ON PLC
    TASK task0(INTERVAL := T#20ms,PRIORITY := 0);
    PROGRAM instance0 WITH task0 : program0;
  END_RESOURCE
END_CONFIGURATION

(* ---- 478-SETUP_MONTHS3.ST ---- *)
TYPE
  oscat_ELEMENT_MONTHS3	: ARRAY [1..12] OF STRING;
  oscat_MONTHS3			: ARRAY [1..3]  OF oscat_ELEMENT_MONTHS3 := [0,0,0];
END_TYPE

FUNCTION_BLOCK SETUP_MONTHS3

	VAR_IN_OUT
		MONTHS3 :	oscat_MONTHS3;
	END_VAR

	VAR
		init :	BOOL;
	END_VAR

	IF init THEN RETURN; END_IF;
	init := TRUE;

	(* ---- english --- *)
	MONTHS3[1][01] := 'Jan';
	MONTHS3[1][02] := 'Feb';
	MONTHS3[1][03] := 'Mar';
	MONTHS3[1][04] := 'Apr';
	MONTHS3[1][05] := 'May';
	MONTHS3[1][06] := 'Jun';
	MONTHS3[1][07] := 'Jul';
	MONTHS3[1][08] := 'Aug';
	MONTHS3[1][09] := 'Sep';
	MONTHS3[1][10] := 'Oct';
	MONTHS3[1][11] := 'Nov';
	MONTHS3[1][12] := 'Dec';

	(* ---- german --- *)
	MONTHS3[2][01] := 'Jan';
	MONTHS3[2][02] := 'Feb';
	MONTHS3[2][03] := 'Mrz';
	MONTHS3[2][04] := 'Apr';
	MONTHs3[2][05] := 'Mai';
	MONTHS3[2][06] := 'Jun';
	MONTHS3[2][07] := 'Jul';
	MONTHS3[2][08] := 'Aug';
	MONTHS3[2][09] := 'Sep';
	MONTHS3[2][10] := 'Okt';
	MONTHS3[2][11] := 'Nov';
	MONTHS3[2][12] := 'Dez';

	(* ---- french --- *)
	MONTHS3[3][01] := 'Jan';
	MONTHS3[3][02] := 'Fev';
	MONTHS3[3][03] := 'Mar';
	MONTHS3[3][04] := 'Avr';
	MONTHs3[3][05] := 'Mai';
	MONTHS3[3][06] := 'Jun';
	MONTHS3[3][07] := 'Jul';
	MONTHS3[3][08] := 'Aou';
	MONTHS3[3][09] := 'Sep';
	MONTHS3[3][10] := 'Oct';
	MONTHS3[3][11] := 'Nov';
	MONTHS3[3][12] := 'Dec';
	(*@KEY@: END_WORKSHEET *)
	END_FUNCTION_BLOCK

PROGRAM program0
  VAR
    LocalVar0 : oscat_MONTHS3;
	func_block : SETUP_MONTHS3;
  END_VAR
	func_block.MONTHS3  := LocalVar0;
	func_block();
	LocalVar0 := func_block.MONTHS3;
END_PROGRAM

CONFIGURATION Config0
  RESOURCE Res0 ON PLC
    TASK task0(INTERVAL := T#20ms,PRIORITY := 0);
    PROGRAM instance0 WITH task0 : program0;
  END_RESOURCE
END_CONFIGURATION
